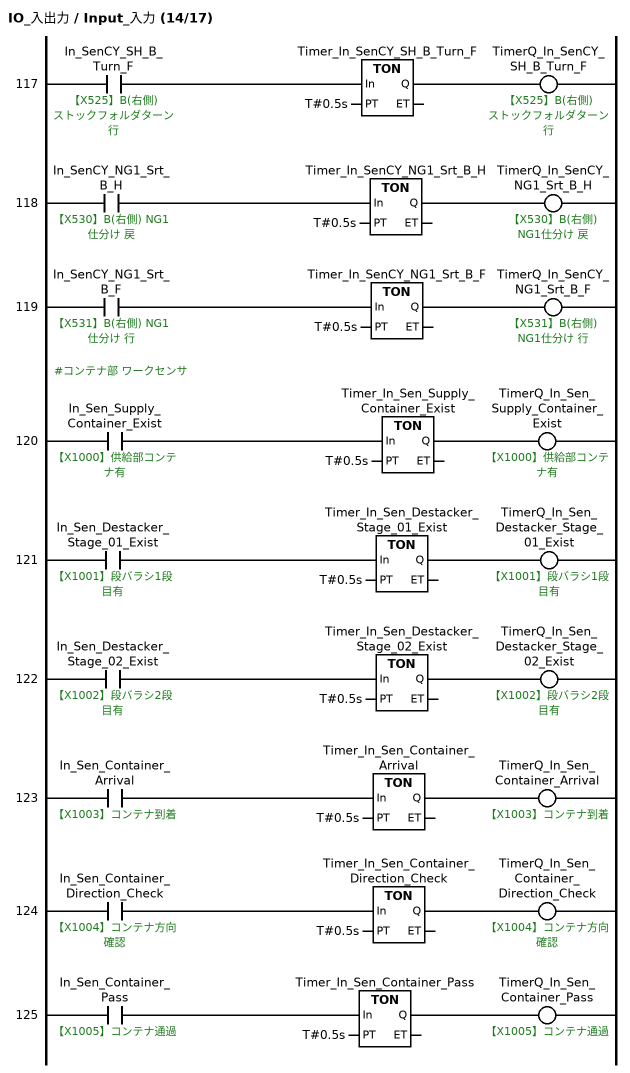
(* [picture p140: IO_入出力 / Input_入力, rungs 117-125] *)
(* Rung 117 *)
Timer_In_SenCY_SH_B_Turn_F(In := In_SenCY_SH_B_Turn_F, PT := T#0.5s);
TimerQ_In_SenCY_SH_B_Turn_F := Timer_In_SenCY_SH_B_Turn_F.Q;
(* Rung 118 *)
Timer_In_SenCY_NG1_Srt_B_H(In := In_SenCY_NG1_Srt_B_H, PT := T#0.5s);
TimerQ_In_SenCY_NG1_Srt_B_H := Timer_In_SenCY_NG1_Srt_B_H.Q;
(* Rung 119 *)
Timer_In_SenCY_NG1_Srt_B_F(In := In_SenCY_NG1_Srt_B_F, PT := T#0.5s);
TimerQ_In_SenCY_NG1_Srt_B_F := Timer_In_SenCY_NG1_Srt_B_F.Q;
(* Rung 120: #コンテナ部 ワークセンサ *)
Timer_In_Sen_Supply_Container_Exist(In := In_Sen_Supply_Container_Exist, PT := T#0.5s);
TimerQ_In_Sen_Supply_Container_Exist := Timer_In_Sen_Supply_Container_Exist.Q;
(* Rung 121 *)
Timer_In_Sen_Destacker_Stage_01_Exist(In := In_Sen_Destacker_Stage_01_Exist, PT := T#0.5s);
TimerQ_In_Sen_Destacker_Stage_01_Exist := Timer_In_Sen_Destacker_Stage_01_Exist.Q;
(* Rung 122 *)
Timer_In_Sen_Destacker_Stage_02_Exist(In := In_Sen_Destacker_Stage_02_Exist, PT := T#0.5s);
TimerQ_In_Sen_Destacker_Stage_02_Exist := Timer_In_Sen_Destacker_Stage_02_Exist.Q;
(* Rung 123 *)
Timer_In_Sen_Container_Arrival(In := In_Sen_Container_Arrival, PT := T#0.5s);
TimerQ_In_Sen_Container_Arrival := Timer_In_Sen_Container_Arrival.Q;
(* Rung 124 *)
Timer_In_Sen_Container_Direction_Check(In := In_Sen_Container_Direction_Check, PT := T#0.5s);
TimerQ_In_Sen_Container_Direction_Check := Timer_In_Sen_Container_Direction_Check.Q;
(* Rung 125 *)
Timer_In_Sen_Container_Pass(In := In_Sen_Container_Pass, PT := T#0.5s);
TimerQ_In_Sen_Container_Pass := Timer_In_Sen_Container_Pass.Q;

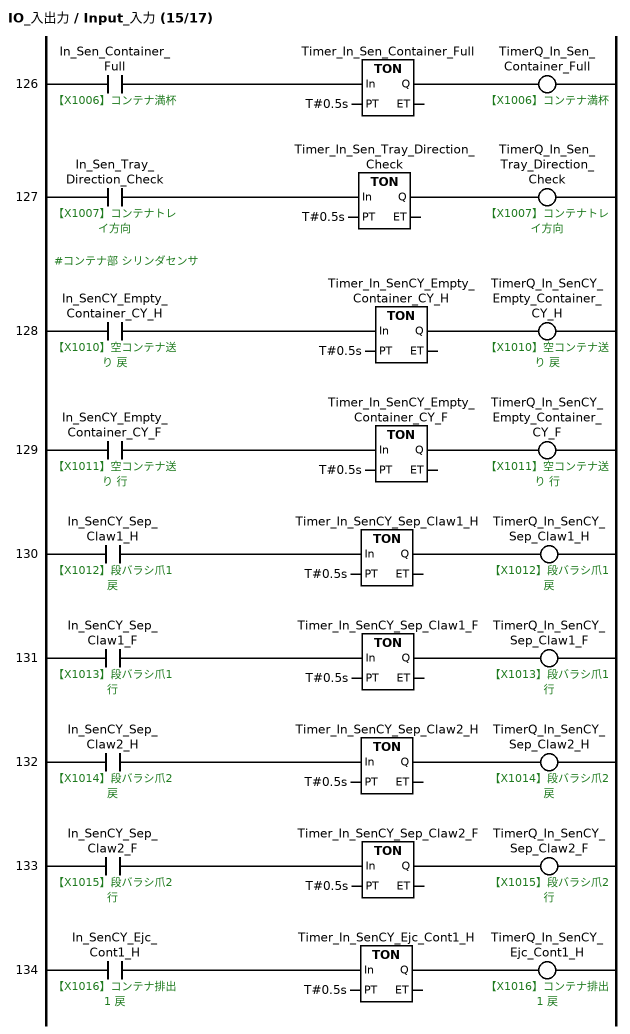
(* Rung 126 *)
Timer_In_Sen_Container_Full(In := In_Sen_Container_Full, PT := T#0.5s);
TimerQ_In_Sen_Container_Full := Timer_In_Sen_Container_Full.Q;
(* Rung 127 *)
Timer_In_Sen_Tray_Direction_Check(In := In_Sen_Tray_Direction_Check, PT := T#0.5s);
TimerQ_In_Sen_Tray_Direction_Check := Timer_In_Sen_Tray_Direction_Check.Q;
(* Rung 128: #コンテナ部 シリンダセンサ *)
Timer_In_SenCY_Empty_Container_CY_H(In := In_SenCY_Empty_Container_CY_H, PT := T#0.5s);
TimerQ_In_SenCY_Empty_Container_CY_H := Timer_In_SenCY_Empty_Container_CY_H.Q;
(* Rung 129 *)
Timer_In_SenCY_Empty_Container_CY_F(In := In_SenCY_Empty_Container_CY_F, PT := T#0.5s);
TimerQ_In_SenCY_Empty_Container_CY_F := Timer_In_SenCY_Empty_Container_CY_F.Q;
(* Rung 130 *)
Timer_In_SenCY_Sep_Claw1_H(In := In_SenCY_Sep_Claw1_H, PT := T#0.5s);
TimerQ_In_SenCY_Sep_Claw1_H := Timer_In_SenCY_Sep_Claw1_H.Q;
(* Rung 131 *)
Timer_In_SenCY_Sep_Claw1_F(In := In_SenCY_Sep_Claw1_F, PT := T#0.5s);
TimerQ_In_SenCY_Sep_Claw1_F := Timer_In_SenCY_Sep_Claw1_F.Q;
(* Rung 132 *)
Timer_In_SenCY_Sep_Claw2_H(In := In_SenCY_Sep_Claw2_H, PT := T#0.5s);
TimerQ_In_SenCY_Sep_Claw2_H := Timer_In_SenCY_Sep_Claw2_H.Q;
(* Rung 133 *)
Timer_In_SenCY_Sep_Claw2_F(In := In_SenCY_Sep_Claw2_F, PT := T#0.5s);
TimerQ_In_SenCY_Sep_Claw2_F := Timer_In_SenCY_Sep_Claw2_F.Q;
(* Rung 134 *)
Timer_In_SenCY_Ejc_Cont1_H(In := In_SenCY_Ejc_Cont1_H, PT := T#0.5s);
TimerQ_In_SenCY_Ejc_Cont1_H := Timer_In_SenCY_Ejc_Cont1_H.Q;

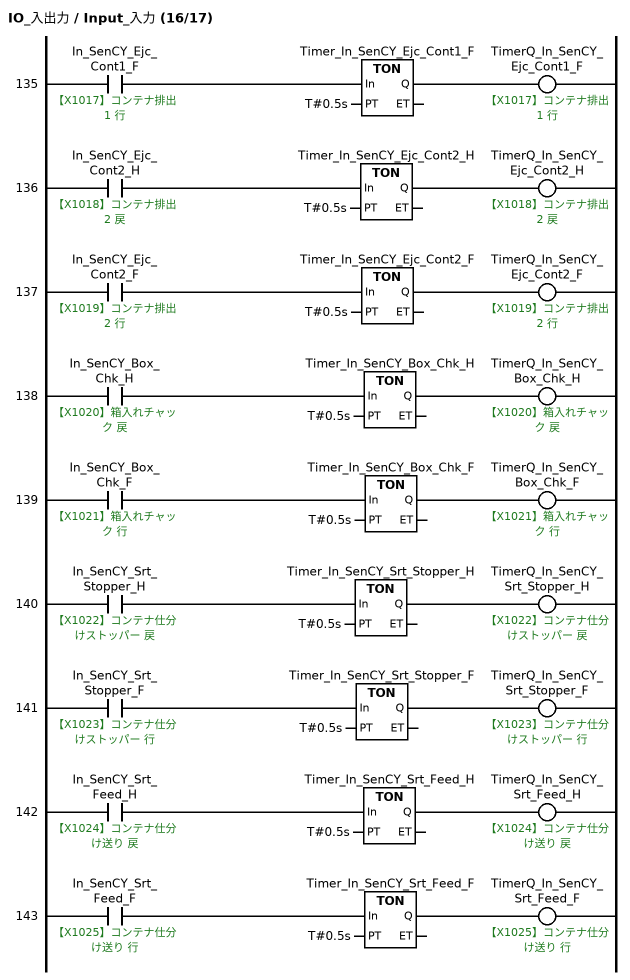
(* Rung 135 *)
Timer_In_SenCY_Ejc_Cont1_F(In := In_SenCY_Ejc_Cont1_F, PT := T#0.5s);
TimerQ_In_SenCY_Ejc_Cont1_F := Timer_In_SenCY_Ejc_Cont1_F.Q;
(* Rung 136 *)
Timer_In_SenCY_Ejc_Cont2_H(In := In_SenCY_Ejc_Cont2_H, PT := T#0.5s);
TimerQ_In_SenCY_Ejc_Cont2_H := Timer_In_SenCY_Ejc_Cont2_H.Q;
(* Rung 137 *)
Timer_In_SenCY_Ejc_Cont2_F(In := In_SenCY_Ejc_Cont2_F, PT := T#0.5s);
TimerQ_In_SenCY_Ejc_Cont2_F := Timer_In_SenCY_Ejc_Cont2_F.Q;
(* Rung 138 *)
Timer_In_SenCY_Box_Chk_H(In := In_SenCY_Box_Chk_H, PT := T#0.5s);
TimerQ_In_SenCY_Box_Chk_H := Timer_In_SenCY_Box_Chk_H.Q;
(* Rung 139 *)
Timer_In_SenCY_Box_Chk_F(In := In_SenCY_Box_Chk_F, PT := T#0.5s);
TimerQ_In_SenCY_Box_Chk_F := Timer_In_SenCY_Box_Chk_F.Q;
(* Rung 140 *)
Timer_In_SenCY_Srt_Stopper_H(In := In_SenCY_Srt_Stopper_H, PT := T#0.5s);
TimerQ_In_SenCY_Srt_Stopper_H := Timer_In_SenCY_Srt_Stopper_H.Q;
(* Rung 141 *)
Timer_In_SenCY_Srt_Stopper_F(In := In_SenCY_Srt_Stopper_F, PT := T#0.5s);
TimerQ_In_SenCY_Srt_Stopper_F := Timer_In_SenCY_Srt_Stopper_F.Q;
(* Rung 142 *)
Timer_In_SenCY_Srt_Feed_H(In := In_SenCY_Srt_Feed_H, PT := T#0.5s);
TimerQ_In_SenCY_Srt_Feed_H := Timer_In_SenCY_Srt_Feed_H.Q;
(* Rung 143 *)
Timer_In_SenCY_Srt_Feed_F(In := In_SenCY_Srt_Feed_F, PT := T#0.5s);
TimerQ_In_SenCY_Srt_Feed_F := Timer_In_SenCY_Srt_Feed_F.Q;

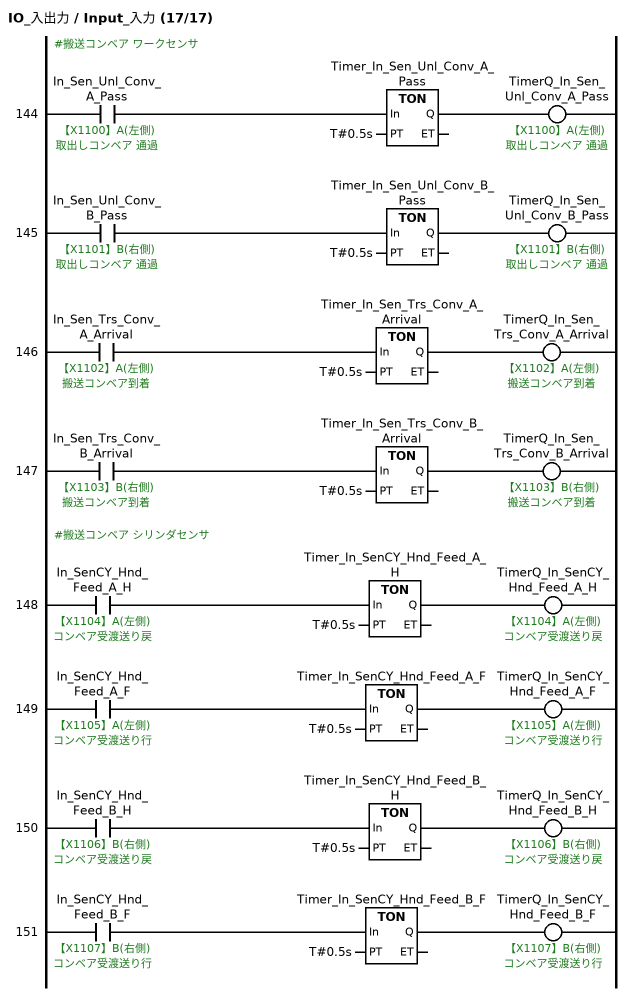
(* Rung 144: #搬送コンベア ワークセンサ *)
Timer_In_Sen_Unl_Conv_A_Pass(In := In_Sen_Unl_Conv_A_Pass, PT := T#0.5s);
TimerQ_In_Sen_Unl_Conv_A_Pass := Timer_In_Sen_Unl_Conv_A_Pass.Q;
(* Rung 145 *)
Timer_In_Sen_Unl_Conv_B_Pass(In := In_Sen_Unl_Conv_B_Pass, PT := T#0.5s);
TimerQ_In_Sen_Unl_Conv_B_Pass := Timer_In_Sen_Unl_Conv_B_Pass.Q;
(* Rung 146 *)
Timer_In_Sen_Trs_Conv_A_Arrival(In := In_Sen_Trs_Conv_A_Arrival, PT := T#0.5s);
TimerQ_In_Sen_Trs_Conv_A_Arrival := Timer_In_Sen_Trs_Conv_A_Arrival.Q;
(* Rung 147 *)
Timer_In_Sen_Trs_Conv_B_Arrival(In := In_Sen_Trs_Conv_B_Arrival, PT := T#0.5s);
TimerQ_In_Sen_Trs_Conv_B_Arrival := Timer_In_Sen_Trs_Conv_B_Arrival.Q;
(* Rung 148: #搬送コンベア シリンダセンサ *)
Timer_In_SenCY_Hnd_Feed_A_H(In := In_SenCY_Hnd_Feed_A_H, PT := T#0.5s);
TimerQ_In_SenCY_Hnd_Feed_A_H := Timer_In_SenCY_Hnd_Feed_A_H.Q;
(* Rung 149 *)
Timer_In_SenCY_Hnd_Feed_A_F(In := In_SenCY_Hnd_Feed_A_F, PT := T#0.5s);
TimerQ_In_SenCY_Hnd_Feed_A_F := Timer_In_SenCY_Hnd_Feed_A_F.Q;
(* Rung 150 *)
Timer_In_SenCY_Hnd_Feed_B_H(In := In_SenCY_Hnd_Feed_B_H, PT := T#0.5s);
TimerQ_In_SenCY_Hnd_Feed_B_H := Timer_In_SenCY_Hnd_Feed_B_H.Q;
(* Rung 151 *)
Timer_In_SenCY_Hnd_Feed_B_F(In := In_SenCY_Hnd_Feed_B_F, PT := T#0.5s);
TimerQ_In_SenCY_Hnd_Feed_B_F := Timer_In_SenCY_Hnd_Feed_B_F.Q;

(* Section Output_出力: ladder, written here as Structured Text *)

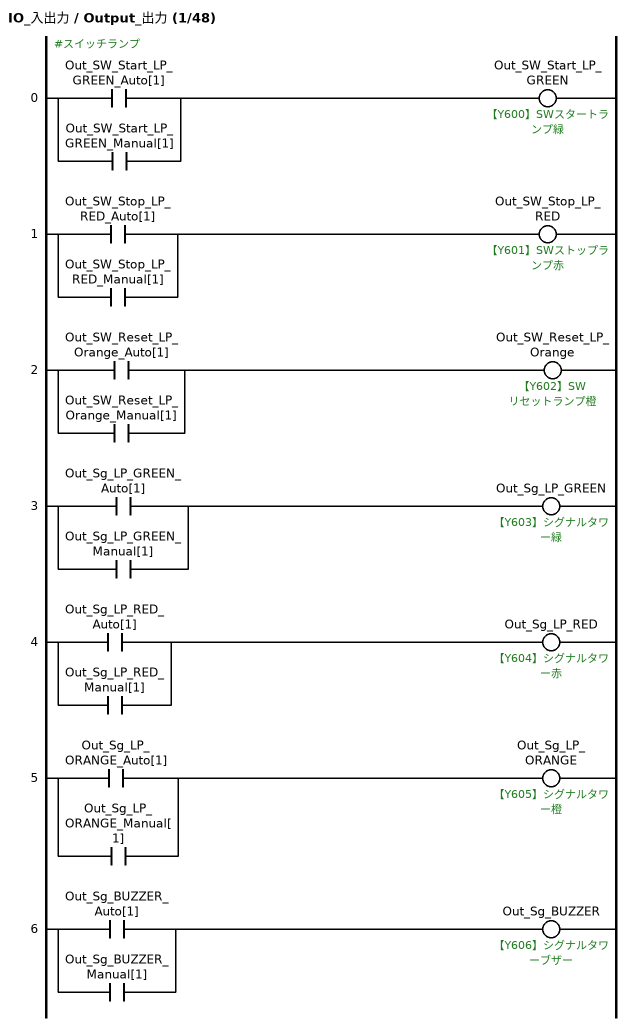
(* Rung 0: #スイッチランプ *)
Out_SW_Start_LP_GREEN := Out_SW_Start_LP_GREEN_Auto[1] OR Out_SW_Start_LP_GREEN_Manual[1];
(* Rung 1 *)
Out_SW_Stop_LP_RED := Out_SW_Stop_LP_RED_Auto[1] OR Out_SW_Stop_LP_RED_Manual[1];
(* Rung 2 *)
Out_SW_Reset_LP_Orange := Out_SW_Reset_LP_Orange_Auto[1] OR Out_SW_Reset_LP_Orange_Manual[1];
(* Rung 3 *)
Out_Sg_LP_GREEN := Out_Sg_LP_GREEN_Auto[1] OR Out_Sg_LP_GREEN_Manual[1];
(* Rung 4 *)
Out_Sg_LP_RED := Out_Sg_LP_RED_Auto[1] OR Out_Sg_LP_RED_Manual[1];
(* Rung 5 *)
Out_Sg_LP_ORANGE := Out_Sg_LP_ORANGE_Auto[1] OR Out_Sg_LP_ORANGE_Manual[1];
(* Rung 6 *)
Out_Sg_BUZZER := Out_Sg_BUZZER_Auto[1] OR Out_Sg_BUZZER_Manual[1];

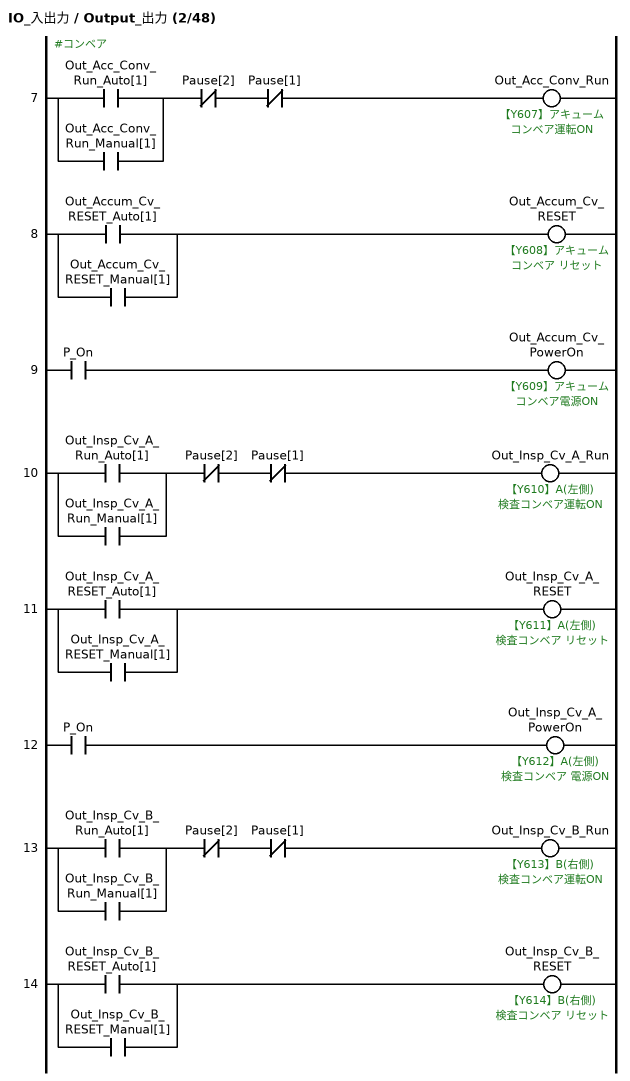
(* Rung 7: #コンベア *)
Out_Acc_Conv_Run := (Out_Acc_Conv_Run_Auto[1] OR Out_Acc_Conv_Run_Manual[1]) AND NOT Pause[2] AND NOT Pause[1];
(* Rung 8 *)
Out_Accum_Cv_RESET := Out_Accum_Cv_RESET_Auto[1] OR Out_Accum_Cv_RESET_Manual[1];
(* Rung 9 *)
Out_Accum_Cv_PowerOn := P_On;
(* Rung 10 *)
Out_Insp_Cv_A_Run := (Out_Insp_Cv_A_Run_Auto[1] OR Out_Insp_Cv_A_Run_Manual[1]) AND NOT Pause[2] AND NOT Pause[1];
(* Rung 11 *)
Out_Insp_Cv_A_RESET := Out_Insp_Cv_A_RESET_Auto[1] OR Out_Insp_Cv_A_RESET_Manual[1];
(* Rung 12 *)
Out_Insp_Cv_A_PowerOn := P_On;
(* Rung 13 *)
Out_Insp_Cv_B_Run := (Out_Insp_Cv_B_Run_Auto[1] OR Out_Insp_Cv_B_Run_Manual[1]) AND NOT Pause[2] AND NOT Pause[1];
(* Rung 14 *)
Out_Insp_Cv_B_RESET := Out_Insp_Cv_B_RESET_Auto[1] OR Out_Insp_Cv_B_RESET_Manual[1];

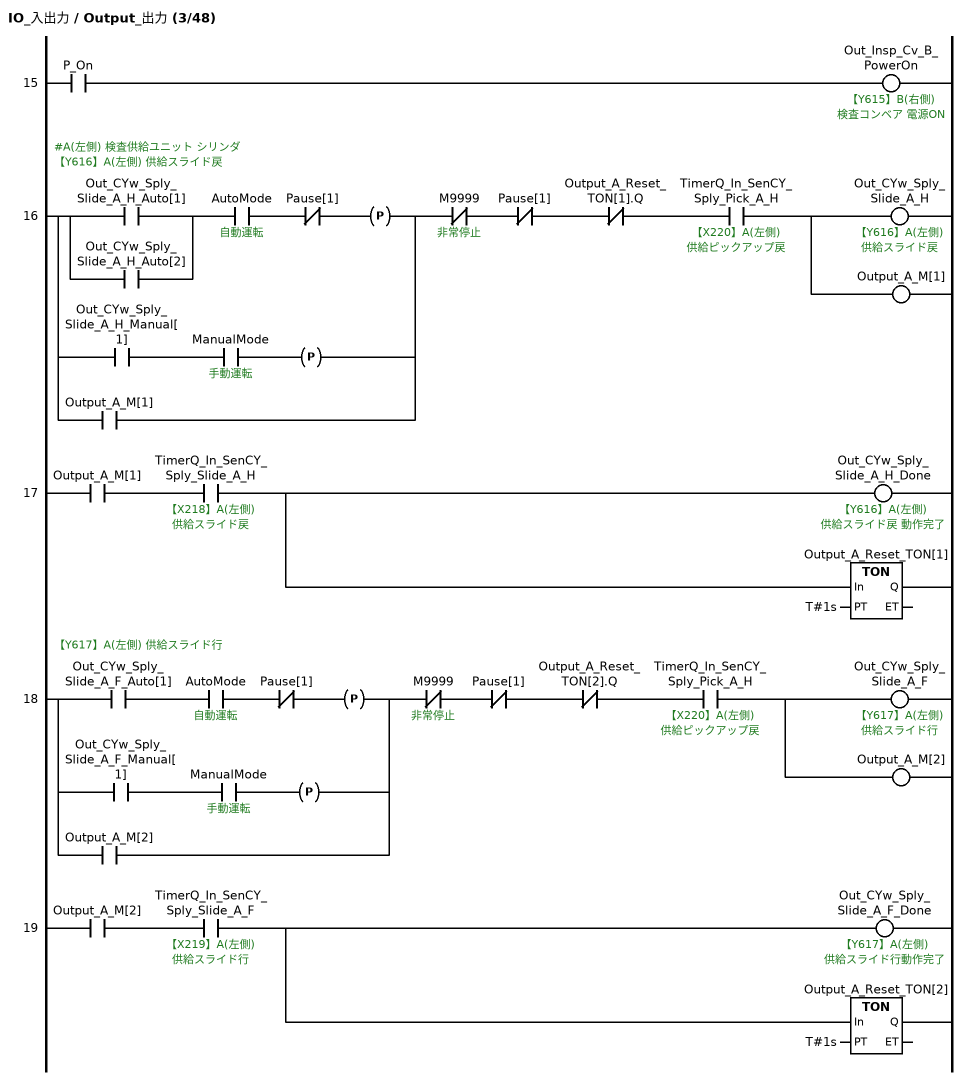
(* Rung 15 *)
Out_Insp_Cv_B_PowerOn := P_On;
(* Rung 16: #A(左側) 検査供給ユニット シリンダ / 【Y616】A(左側) 供給スライド戻 *)
_e1(CLK := (Out_CYw_Sply_Slide_A_H_Auto[1] OR Out_CYw_Sply_Slide_A_H_Auto[2]) AND AutoMode AND NOT Pause[1]);
_e2(CLK := Out_CYw_Sply_Slide_A_H_Manual[1] AND ManualMode);
_p3 := (_e1.Q OR _e2.Q OR Output_A_M[1]) AND NOT M9999 AND NOT Pause[1] AND NOT Output_A_Reset_TON[1].Q AND TimerQ_In_SenCY_Sply_Pick_A_H;
Out_CYw_Sply_Slide_A_H := _p3;
Output_A_M[1] := _p3;
(* Rung 17 *)
Out_CYw_Sply_Slide_A_H_Done := Output_A_M[1] AND TimerQ_In_SenCY_Sply_Slide_A_H;
Output_A_Reset_TON[1](In := Output_A_M[1] AND TimerQ_In_SenCY_Sply_Slide_A_H, PT := T#1s);
(* Rung 18: 【Y617】A(左側) 供給スライド行 *)
_e4(CLK := Out_CYw_Sply_Slide_A_F_Auto[1] AND AutoMode AND NOT Pause[1]);
_e5(CLK := Out_CYw_Sply_Slide_A_F_Manual[1] AND ManualMode);
_p6 := (_e4.Q OR _e5.Q OR Output_A_M[2]) AND NOT M9999 AND NOT Pause[1] AND NOT Output_A_Reset_TON[2].Q AND TimerQ_In_SenCY_Sply_Pick_A_H;
Out_CYw_Sply_Slide_A_F := _p6;
Output_A_M[2] := _p6;
(* Rung 19 *)
Out_CYw_Sply_Slide_A_F_Done := Output_A_M[2] AND TimerQ_In_SenCY_Sply_Slide_A_F;
Output_A_Reset_TON[2](In := Output_A_M[2] AND TimerQ_In_SenCY_Sply_Slide_A_F, PT := T#1s);

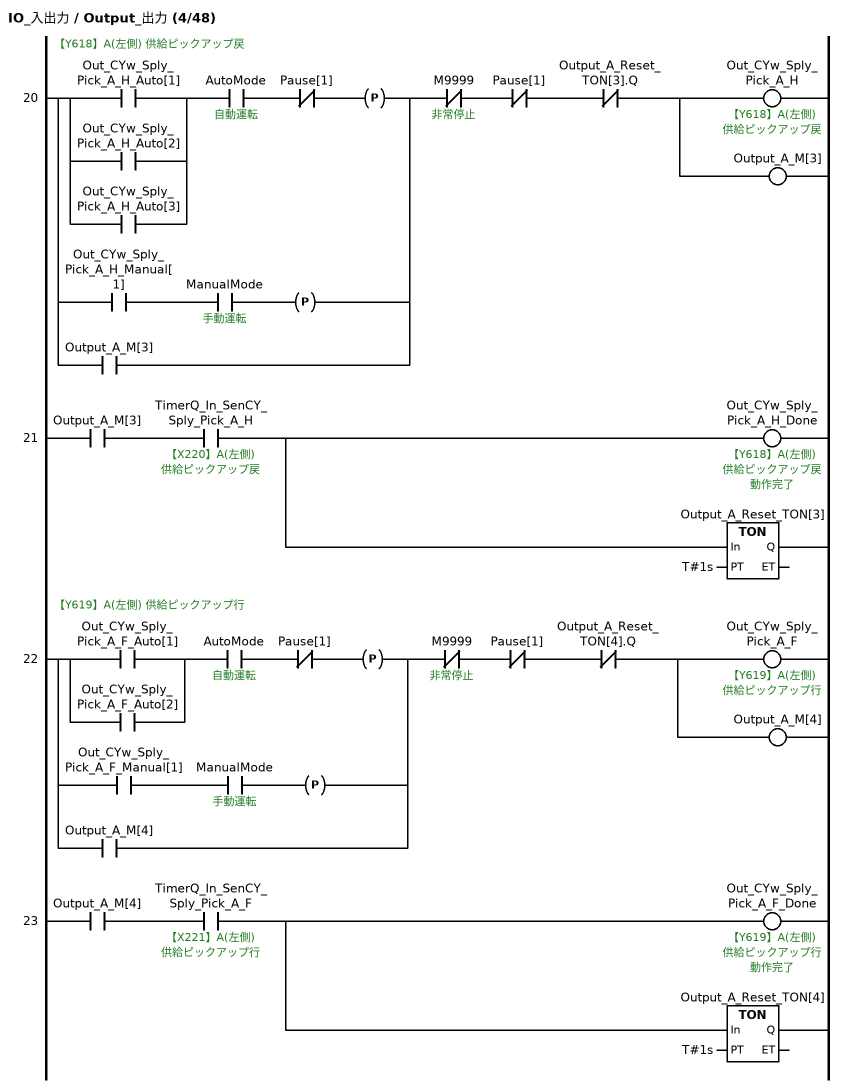
(* Rung 20: 【Y618】A(左側) 供給ピックアップ戻 *)
_e7(CLK := (Out_CYw_Sply_Pick_A_H_Auto[1] OR Out_CYw_Sply_Pick_A_H_Auto[2] OR Out_CYw_Sply_Pick_A_H_Auto[3]) AND AutoMode AND NOT Pause[1]);
_e8(CLK := Out_CYw_Sply_Pick_A_H_Manual[1] AND ManualMode);
_p9 := (_e7.Q OR _e8.Q OR Output_A_M[3]) AND NOT M9999 AND NOT Pause[1] AND NOT Output_A_Reset_TON[3].Q;
Out_CYw_Sply_Pick_A_H := _p9;
Output_A_M[3] := _p9;
(* Rung 21 *)
Out_CYw_Sply_Pick_A_H_Done := Output_A_M[3] AND TimerQ_In_SenCY_Sply_Pick_A_H;
Output_A_Reset_TON[3](In := Output_A_M[3] AND TimerQ_In_SenCY_Sply_Pick_A_H, PT := T#1s);
(* Rung 22: 【Y619】A(左側) 供給ピックアップ行 *)
_e10(CLK := (Out_CYw_Sply_Pick_A_F_Auto[1] OR Out_CYw_Sply_Pick_A_F_Auto[2]) AND AutoMode AND NOT Pause[1]);
_e11(CLK := Out_CYw_Sply_Pick_A_F_Manual[1] AND ManualMode);
_p12 := (_e10.Q OR _e11.Q OR Output_A_M[4]) AND NOT M9999 AND NOT Pause[1] AND NOT Output_A_Reset_TON[4].Q;
Out_CYw_Sply_Pick_A_F := _p12;
Output_A_M[4] := _p12;
(* Rung 23 *)
Out_CYw_Sply_Pick_A_F_Done := Output_A_M[4] AND TimerQ_In_SenCY_Sply_Pick_A_F;
Output_A_Reset_TON[4](In := Output_A_M[4] AND TimerQ_In_SenCY_Sply_Pick_A_F, PT := T#1s);

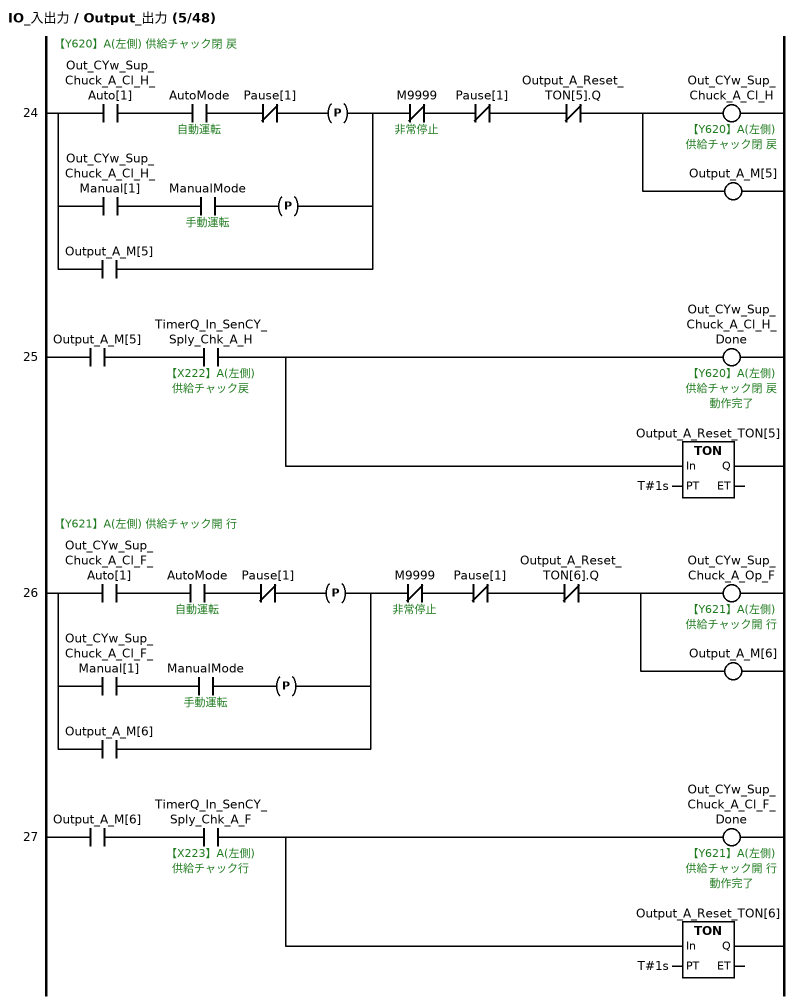
(* Rung 24: 【Y620】A(左側) 供給チャック閉 戻 *)
_e13(CLK := Out_CYw_Sup_Chuck_A_Cl_H_Auto[1] AND AutoMode AND NOT Pause[1]);
_e14(CLK := Out_CYw_Sup_Chuck_A_Cl_H_Manual[1] AND ManualMode);
_p15 := (_e13.Q OR _e14.Q OR Output_A_M[5]) AND NOT M9999 AND NOT Pause[1] AND NOT Output_A_Reset_TON[5].Q;
Out_CYw_Sup_Chuck_A_Cl_H := _p15;
Output_A_M[5] := _p15;
(* Rung 25 *)
Out_CYw_Sup_Chuck_A_Cl_H_Done := Output_A_M[5] AND TimerQ_In_SenCY_Sply_Chk_A_H;
Output_A_Reset_TON[5](In := Output_A_M[5] AND TimerQ_In_SenCY_Sply_Chk_A_H, PT := T#1s);
(* Rung 26: 【Y621】A(左側) 供給チャック開 行 *)
_e16(CLK := Out_CYw_Sup_Chuck_A_Cl_F_Auto[1] AND AutoMode AND NOT Pause[1]);
_e17(CLK := Out_CYw_Sup_Chuck_A_Cl_F_Manual[1] AND ManualMode);
_p18 := (_e16.Q OR _e17.Q OR Output_A_M[6]) AND NOT M9999 AND NOT Pause[1] AND NOT Output_A_Reset_TON[6].Q;
Out_CYw_Sup_Chuck_A_Op_F := _p18;
Output_A_M[6] := _p18;
(* Rung 27 *)
Out_CYw_Sup_Chuck_A_Cl_F_Done := Output_A_M[6] AND TimerQ_In_SenCY_Sply_Chk_A_F;
Output_A_Reset_TON[6](In := Output_A_M[6] AND TimerQ_In_SenCY_Sply_Chk_A_F, PT := T#1s);

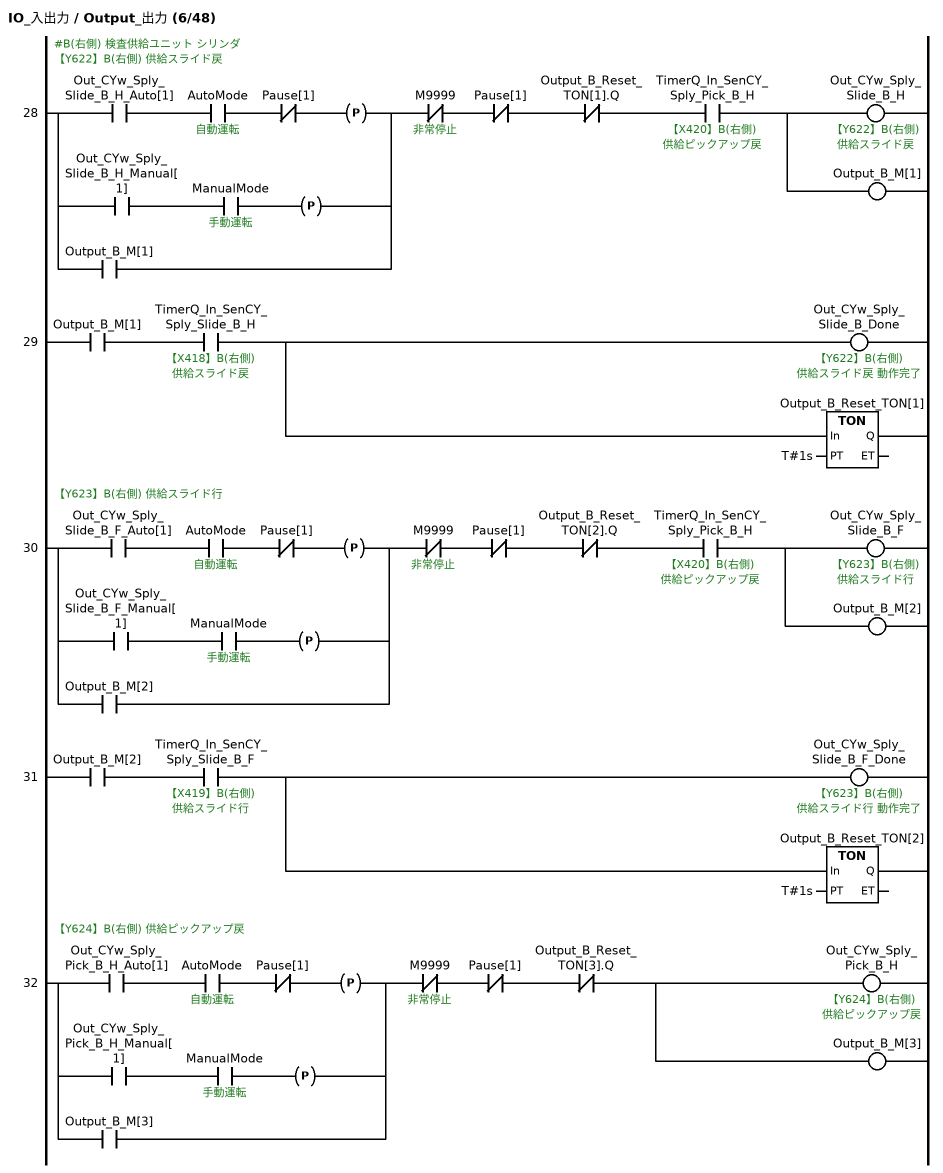
(* Rung 28: #B(右側) 検査供給ユニット シリンダ / 【Y622】B(右側) 供給スライド戻 *)
_e19(CLK := Out_CYw_Sply_Slide_B_H_Auto[1] AND AutoMode AND NOT Pause[1]);
_e20(CLK := Out_CYw_Sply_Slide_B_H_Manual[1] AND ManualMode);
_p21 := (_e19.Q OR _e20.Q OR Output_B_M[1]) AND NOT M9999 AND NOT Pause[1] AND NOT Output_B_Reset_TON[1].Q AND TimerQ_In_SenCY_Sply_Pick_B_H;
Out_CYw_Sply_Slide_B_H := _p21;
Output_B_M[1] := _p21;
(* Rung 29 *)
Out_CYw_Sply_Slide_B_Done := Output_B_M[1] AND TimerQ_In_SenCY_Sply_Slide_B_H;
Output_B_Reset_TON[1](In := Output_B_M[1] AND TimerQ_In_SenCY_Sply_Slide_B_H, PT := T#1s);
(* Rung 30: 【Y623】B(右側) 供給スライド行 *)
_e22(CLK := Out_CYw_Sply_Slide_B_F_Auto[1] AND AutoMode AND NOT Pause[1]);
_e23(CLK := Out_CYw_Sply_Slide_B_F_Manual[1] AND ManualMode);
_p24 := (_e22.Q OR _e23.Q OR Output_B_M[2]) AND NOT M9999 AND NOT Pause[1] AND NOT Output_B_Reset_TON[2].Q AND TimerQ_In_SenCY_Sply_Pick_B_H;
Out_CYw_Sply_Slide_B_F := _p24;
Output_B_M[2] := _p24;
(* Rung 31 *)
Out_CYw_Sply_Slide_B_F_Done := Output_B_M[2] AND TimerQ_In_SenCY_Sply_Slide_B_F;
Output_B_Reset_TON[2](In := Output_B_M[2] AND TimerQ_In_SenCY_Sply_Slide_B_F, PT := T#1s);
(* Rung 32: 【Y624】B(右側) 供給ピックアップ戻 *)
_e25(CLK := Out_CYw_Sply_Pick_B_H_Auto[1] AND AutoMode AND NOT Pause[1]);
_e26(CLK := Out_CYw_Sply_Pick_B_H_Manual[1] AND ManualMode);
_p27 := (_e25.Q OR _e26.Q OR Output_B_M[3]) AND NOT M9999 AND NOT Pause[1] AND NOT Output_B_Reset_TON[3].Q;
Out_CYw_Sply_Pick_B_H := _p27;
Output_B_M[3] := _p27;

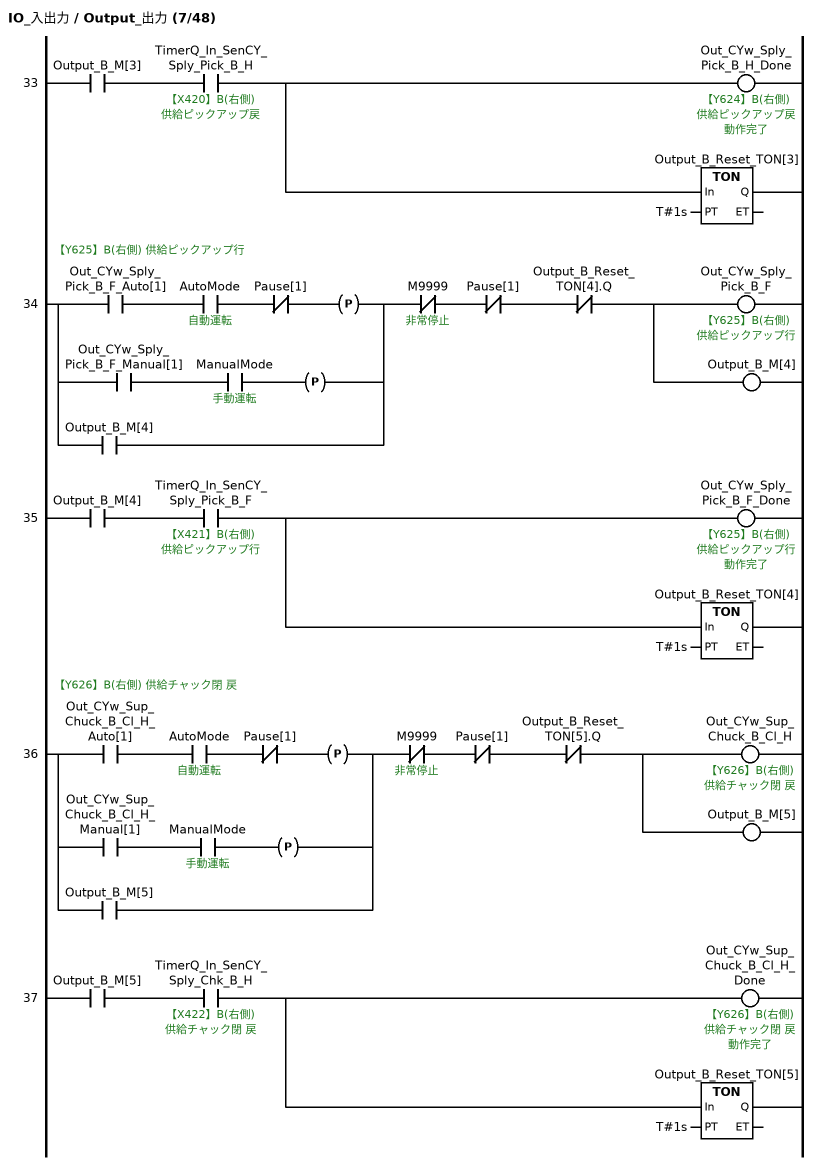
(* Rung 33 *)
Out_CYw_Sply_Pick_B_H_Done := Output_B_M[3] AND TimerQ_In_SenCY_Sply_Pick_B_H;
Output_B_Reset_TON[3](In := Output_B_M[3] AND TimerQ_In_SenCY_Sply_Pick_B_H, PT := T#1s);
(* Rung 34: 【Y625】B(右側) 供給ピックアップ行 *)
_e28(CLK := Out_CYw_Sply_Pick_B_F_Auto[1] AND AutoMode AND NOT Pause[1]);
_e29(CLK := Out_CYw_Sply_Pick_B_F_Manual[1] AND ManualMode);
_p30 := (_e28.Q OR _e29.Q OR Output_B_M[4]) AND NOT M9999 AND NOT Pause[1] AND NOT Output_B_Reset_TON[4].Q;
Out_CYw_Sply_Pick_B_F := _p30;
Output_B_M[4] := _p30;
(* Rung 35 *)
Out_CYw_Sply_Pick_B_F_Done := Output_B_M[4] AND TimerQ_In_SenCY_Sply_Pick_B_F;
Output_B_Reset_TON[4](In := Output_B_M[4] AND TimerQ_In_SenCY_Sply_Pick_B_F, PT := T#1s);
(* Rung 36: 【Y626】B(右側) 供給チャック閉 戻 *)
_e31(CLK := Out_CYw_Sup_Chuck_B_Cl_H_Auto[1] AND AutoMode AND NOT Pause[1]);
_e32(CLK := Out_CYw_Sup_Chuck_B_Cl_H_Manual[1] AND ManualMode);
_p33 := (_e31.Q OR _e32.Q OR Output_B_M[5]) AND NOT M9999 AND NOT Pause[1] AND NOT Output_B_Reset_TON[5].Q;
Out_CYw_Sup_Chuck_B_Cl_H := _p33;
Output_B_M[5] := _p33;
(* Rung 37 *)
Out_CYw_Sup_Chuck_B_Cl_H_Done := Output_B_M[5] AND TimerQ_In_SenCY_Sply_Chk_B_H;
Output_B_Reset_TON[5](In := Output_B_M[5] AND TimerQ_In_SenCY_Sply_Chk_B_H, PT := T#1s);

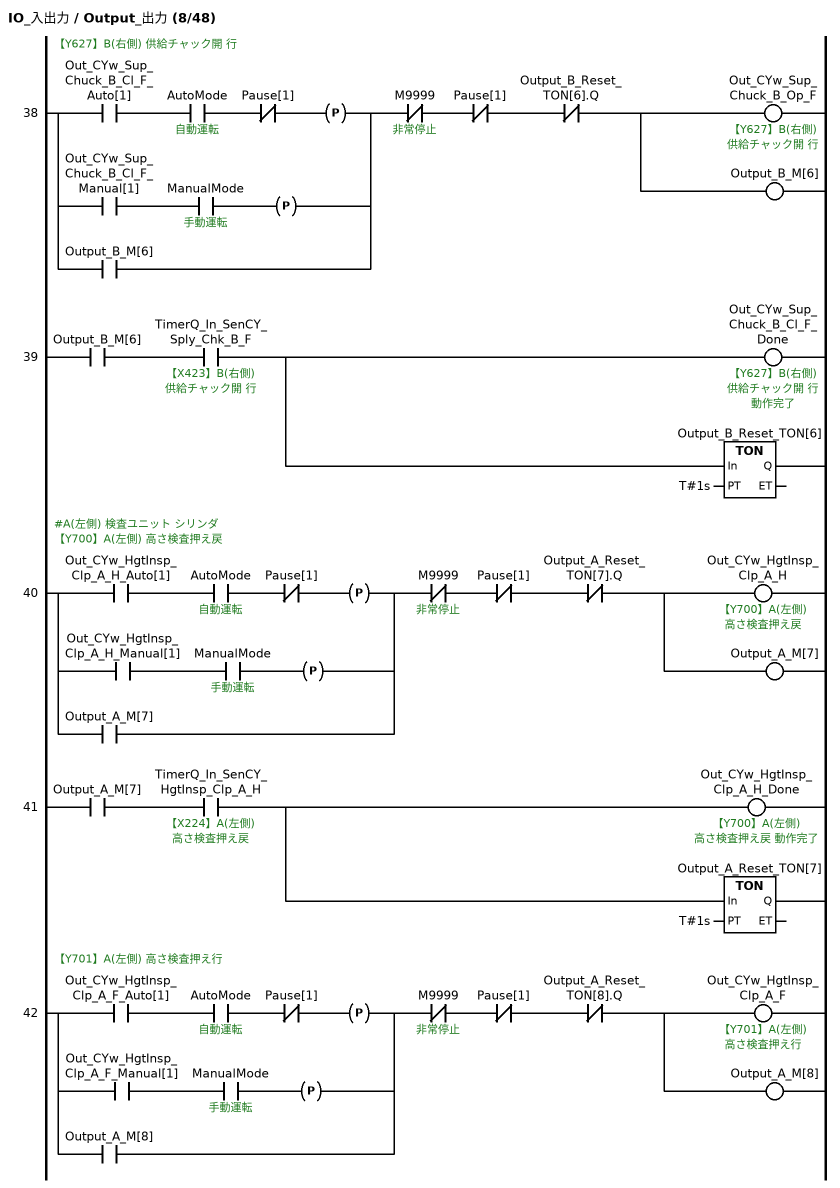
(* Rung 38: 【Y627】B(右側) 供給チャック開 行 *)
_e34(CLK := Out_CYw_Sup_Chuck_B_Cl_F_Auto[1] AND AutoMode AND NOT Pause[1]);
_e35(CLK := Out_CYw_Sup_Chuck_B_Cl_F_Manual[1] AND ManualMode);
_p36 := (_e34.Q OR _e35.Q OR Output_B_M[6]) AND NOT M9999 AND NOT Pause[1] AND NOT Output_B_Reset_TON[6].Q;
Out_CYw_Sup_Chuck_B_Op_F := _p36;
Output_B_M[6] := _p36;
(* Rung 39 *)
Out_CYw_Sup_Chuck_B_Cl_F_Done := Output_B_M[6] AND TimerQ_In_SenCY_Sply_Chk_B_F;
Output_B_Reset_TON[6](In := Output_B_M[6] AND TimerQ_In_SenCY_Sply_Chk_B_F, PT := T#1s);
(* Rung 40: #A(左側) 検査ユニット シリンダ / 【Y700】A(左側) 高さ検査押え戻 *)
_e37(CLK := Out_CYw_HgtInsp_Clp_A_H_Auto[1] AND AutoMode AND NOT Pause[1]);
_e38(CLK := Out_CYw_HgtInsp_Clp_A_H_Manual[1] AND ManualMode);
_p39 := (_e37.Q OR _e38.Q OR Output_A_M[7]) AND NOT M9999 AND NOT Pause[1] AND NOT Output_A_Reset_TON[7].Q;
Out_CYw_HgtInsp_Clp_A_H := _p39;
Output_A_M[7] := _p39;
(* Rung 41 *)
_p40 := Output_A_M[7] AND TimerQ_In_SenCY_HgtInsp_Clp_A_H;
Out_CYw_HgtInsp_Clp_A_H_Done := _p40;
Output_A_Reset_TON[7](In := _p40, PT := T#1s);
(* Rung 42: 【Y701】A(左側) 高さ検査押え行 *)
_e41(CLK := Out_CYw_HgtInsp_Clp_A_F_Auto[1] AND AutoMode AND NOT Pause[1]);
_e42(CLK := Out_CYw_HgtInsp_Clp_A_F_Manual[1] AND ManualMode);
_p43 := (_e41.Q OR _e42.Q OR Output_A_M[8]) AND NOT M9999 AND NOT Pause[1] AND NOT Output_A_Reset_TON[8].Q;
Out_CYw_HgtInsp_Clp_A_F := _p43;
Output_A_M[8] := _p43;

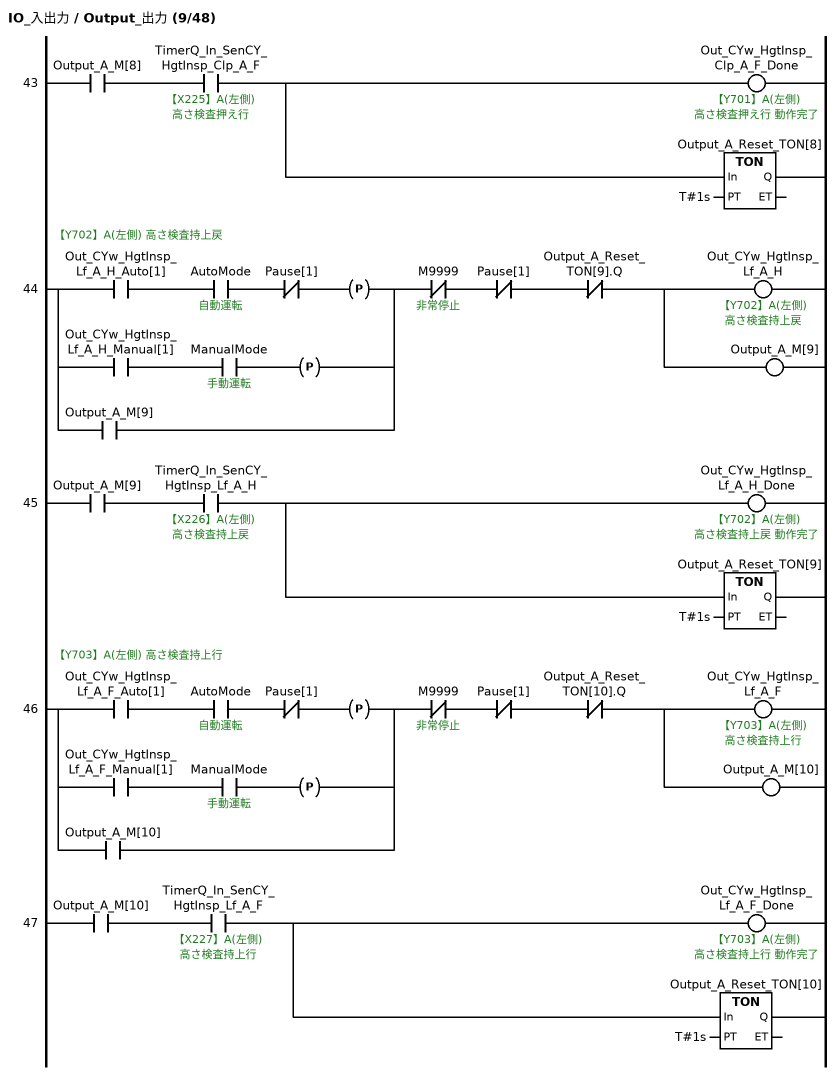
(* Rung 43 *)
_p44 := Output_A_M[8] AND TimerQ_In_SenCY_HgtInsp_Clp_A_F;
Out_CYw_HgtInsp_Clp_A_F_Done := _p44;
Output_A_Reset_TON[8](In := _p44, PT := T#1s);
(* Rung 44: 【Y702】A(左側) 高さ検査持上戻 *)
_e45(CLK := Out_CYw_HgtInsp_Lf_A_H_Auto[1] AND AutoMode AND NOT Pause[1]);
_e46(CLK := Out_CYw_HgtInsp_Lf_A_H_Manual[1] AND ManualMode);
_p47 := (_e45.Q OR _e46.Q OR Output_A_M[9]) AND NOT M9999 AND NOT Pause[1] AND NOT Output_A_Reset_TON[9].Q;
Out_CYw_HgtInsp_Lf_A_H := _p47;
Output_A_M[9] := _p47;
(* Rung 45 *)
Out_CYw_HgtInsp_Lf_A_H_Done := Output_A_M[9] AND TimerQ_In_SenCY_HgtInsp_Lf_A_H;
Output_A_Reset_TON[9](In := Output_A_M[9] AND TimerQ_In_SenCY_HgtInsp_Lf_A_H, PT := T#1s);
(* Rung 46: 【Y703】A(左側) 高さ検査持上行 *)
_e48(CLK := Out_CYw_HgtInsp_Lf_A_F_Auto[1] AND AutoMode AND NOT Pause[1]);
_e49(CLK := Out_CYw_HgtInsp_Lf_A_F_Manual[1] AND ManualMode);
_p50 := (_e48.Q OR _e49.Q OR Output_A_M[10]) AND NOT M9999 AND NOT Pause[1] AND NOT Output_A_Reset_TON[10].Q;
Out_CYw_HgtInsp_Lf_A_F := _p50;
Output_A_M[10] := _p50;
(* Rung 47 *)
_p51 := Output_A_M[10] AND TimerQ_In_SenCY_HgtInsp_Lf_A_F;
Out_CYw_HgtInsp_Lf_A_F_Done := _p51;
Output_A_Reset_TON[10](In := _p51, PT := T#1s);

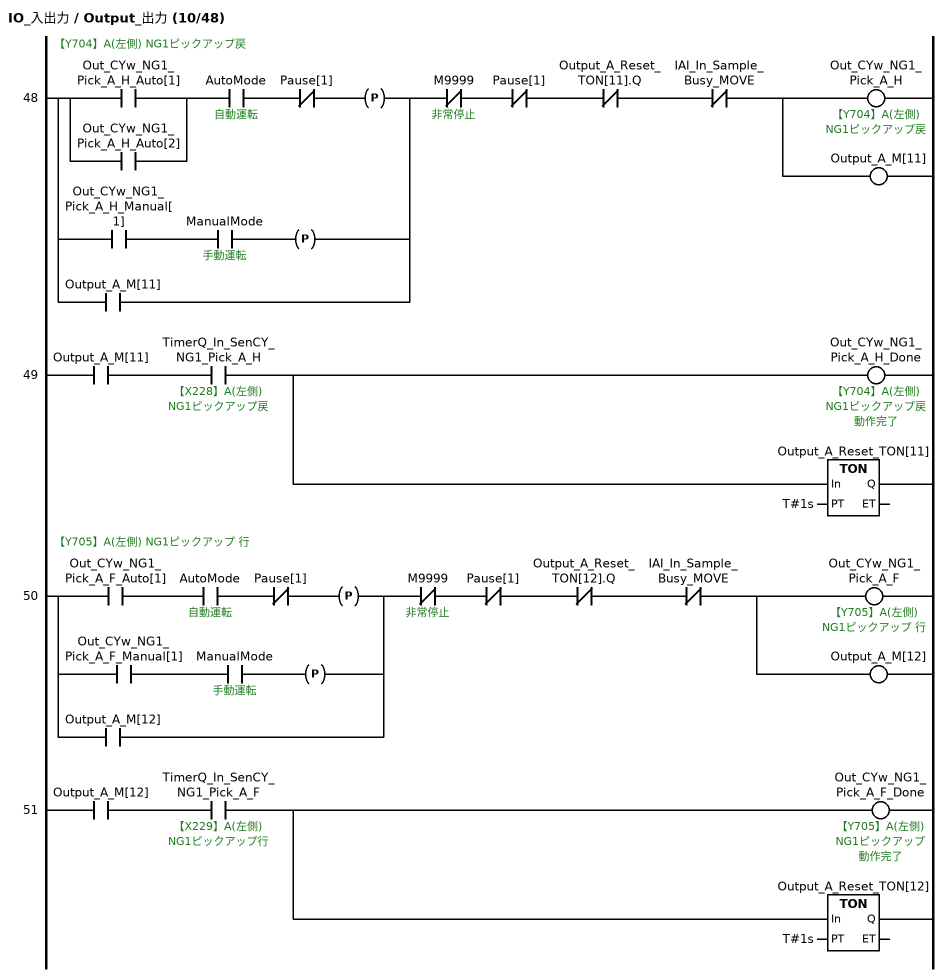
(* Rung 48: 【Y704】A(左側) NG1ピックアップ戻 *)
_e52(CLK := (Out_CYw_NG1_Pick_A_H_Auto[1] OR Out_CYw_NG1_Pick_A_H_Auto[2]) AND AutoMode AND NOT Pause[1]);
_e53(CLK := Out_CYw_NG1_Pick_A_H_Manual[1] AND ManualMode);
_p54 := (_e52.Q OR _e53.Q OR Output_A_M[11]) AND NOT M9999 AND NOT Pause[1] AND NOT Output_A_Reset_TON[11].Q AND NOT IAI_In_Sample_Busy_MOVE;
Out_CYw_NG1_Pick_A_H := _p54;
Output_A_M[11] := _p54;
(* Rung 49 *)
Out_CYw_NG1_Pick_A_H_Done := Output_A_M[11] AND TimerQ_In_SenCY_NG1_Pick_A_H;
Output_A_Reset_TON[11](In := Output_A_M[11] AND TimerQ_In_SenCY_NG1_Pick_A_H, PT := T#1s);
(* Rung 50: 【Y705】A(左側) NG1ピックアップ 行 *)
_e55(CLK := Out_CYw_NG1_Pick_A_F_Auto[1] AND AutoMode AND NOT Pause[1]);
_e56(CLK := Out_CYw_NG1_Pick_A_F_Manual[1] AND ManualMode);
_p57 := (_e55.Q OR _e56.Q OR Output_A_M[12]) AND NOT M9999 AND NOT Pause[1] AND NOT Output_A_Reset_TON[12].Q AND NOT IAI_In_Sample_Busy_MOVE;
Out_CYw_NG1_Pick_A_F := _p57;
Output_A_M[12] := _p57;
(* Rung 51 *)
Out_CYw_NG1_Pick_A_F_Done := Output_A_M[12] AND TimerQ_In_SenCY_NG1_Pick_A_F;
Output_A_Reset_TON[12](In := Output_A_M[12] AND TimerQ_In_SenCY_NG1_Pick_A_F, PT := T#1s);

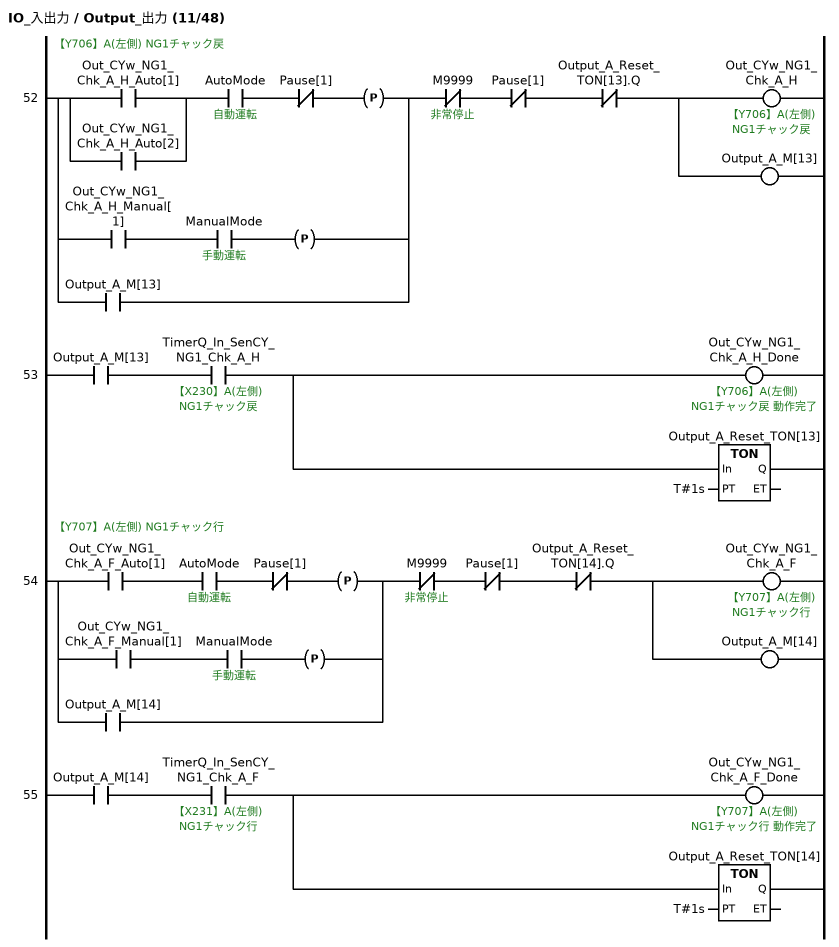
(* Rung 52: 【Y706】A(左側) NG1チャック戻 *)
_e58(CLK := (Out_CYw_NG1_Chk_A_H_Auto[1] OR Out_CYw_NG1_Chk_A_H_Auto[2]) AND AutoMode AND NOT Pause[1]);
_e59(CLK := Out_CYw_NG1_Chk_A_H_Manual[1] AND ManualMode);
_p60 := (_e58.Q OR _e59.Q OR Output_A_M[13]) AND NOT M9999 AND NOT Pause[1] AND NOT Output_A_Reset_TON[13].Q;
Out_CYw_NG1_Chk_A_H := _p60;
Output_A_M[13] := _p60;
(* Rung 53 *)
Out_CYw_NG1_Chk_A_H_Done := Output_A_M[13] AND TimerQ_In_SenCY_NG1_Chk_A_H;
Output_A_Reset_TON[13](In := Output_A_M[13] AND TimerQ_In_SenCY_NG1_Chk_A_H, PT := T#1s);
(* Rung 54: 【Y707】A(左側) NG1チャック行 *)
_e61(CLK := Out_CYw_NG1_Chk_A_F_Auto[1] AND AutoMode AND NOT Pause[1]);
_e62(CLK := Out_CYw_NG1_Chk_A_F_Manual[1] AND ManualMode);
_p63 := (_e61.Q OR _e62.Q OR Output_A_M[14]) AND NOT M9999 AND NOT Pause[1] AND NOT Output_A_Reset_TON[14].Q;
Out_CYw_NG1_Chk_A_F := _p63;
Output_A_M[14] := _p63;
(* Rung 55 *)
Out_CYw_NG1_Chk_A_F_Done := Output_A_M[14] AND TimerQ_In_SenCY_NG1_Chk_A_F;
Output_A_Reset_TON[14](In := Output_A_M[14] AND TimerQ_In_SenCY_NG1_Chk_A_F, PT := T#1s);

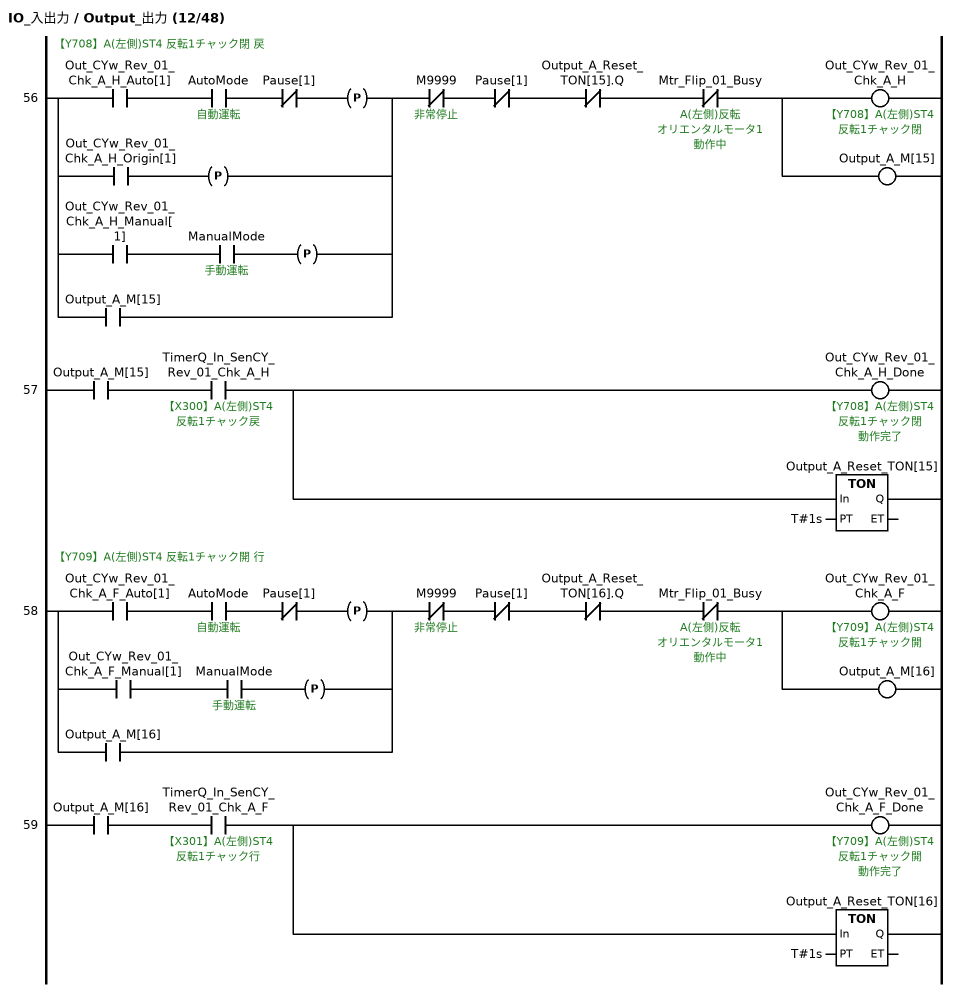
(* Rung 56: 【Y708】A(左側)ST4 反転1チャック閉 戻 *)
_e64(CLK := Out_CYw_Rev_01_Chk_A_H_Auto[1] AND AutoMode AND NOT Pause[1]);
_e65(CLK := Out_CYw_Rev_01_Chk_A_H_Origin[1]);
_e66(CLK := Out_CYw_Rev_01_Chk_A_H_Manual[1] AND ManualMode);
_p67 := (_e64.Q OR _e65.Q OR _e66.Q OR Output_A_M[15]) AND NOT M9999 AND NOT Pause[1] AND NOT Output_A_Reset_TON[15].Q AND NOT Mtr_Flip_01_Busy;
Out_CYw_Rev_01_Chk_A_H := _p67;
Output_A_M[15] := _p67;
(* Rung 57 *)
_p68 := Output_A_M[15] AND TimerQ_In_SenCY_Rev_01_Chk_A_H;
Out_CYw_Rev_01_Chk_A_H_Done := _p68;
Output_A_Reset_TON[15](In := _p68, PT := T#1s);
(* Rung 58: 【Y709】A(左側)ST4 反転1チャック開 行 *)
_e69(CLK := Out_CYw_Rev_01_Chk_A_F_Auto[1] AND AutoMode AND NOT Pause[1]);
_e70(CLK := Out_CYw_Rev_01_Chk_A_F_Manual[1] AND ManualMode);
_p71 := (_e69.Q OR _e70.Q OR Output_A_M[16]) AND NOT M9999 AND NOT Pause[1] AND NOT Output_A_Reset_TON[16].Q AND NOT Mtr_Flip_01_Busy;
Out_CYw_Rev_01_Chk_A_F := _p71;
Output_A_M[16] := _p71;
(* Rung 59 *)
_p72 := Output_A_M[16] AND TimerQ_In_SenCY_Rev_01_Chk_A_F;
Out_CYw_Rev_01_Chk_A_F_Done := _p72;
Output_A_Reset_TON[16](In := _p72, PT := T#1s);

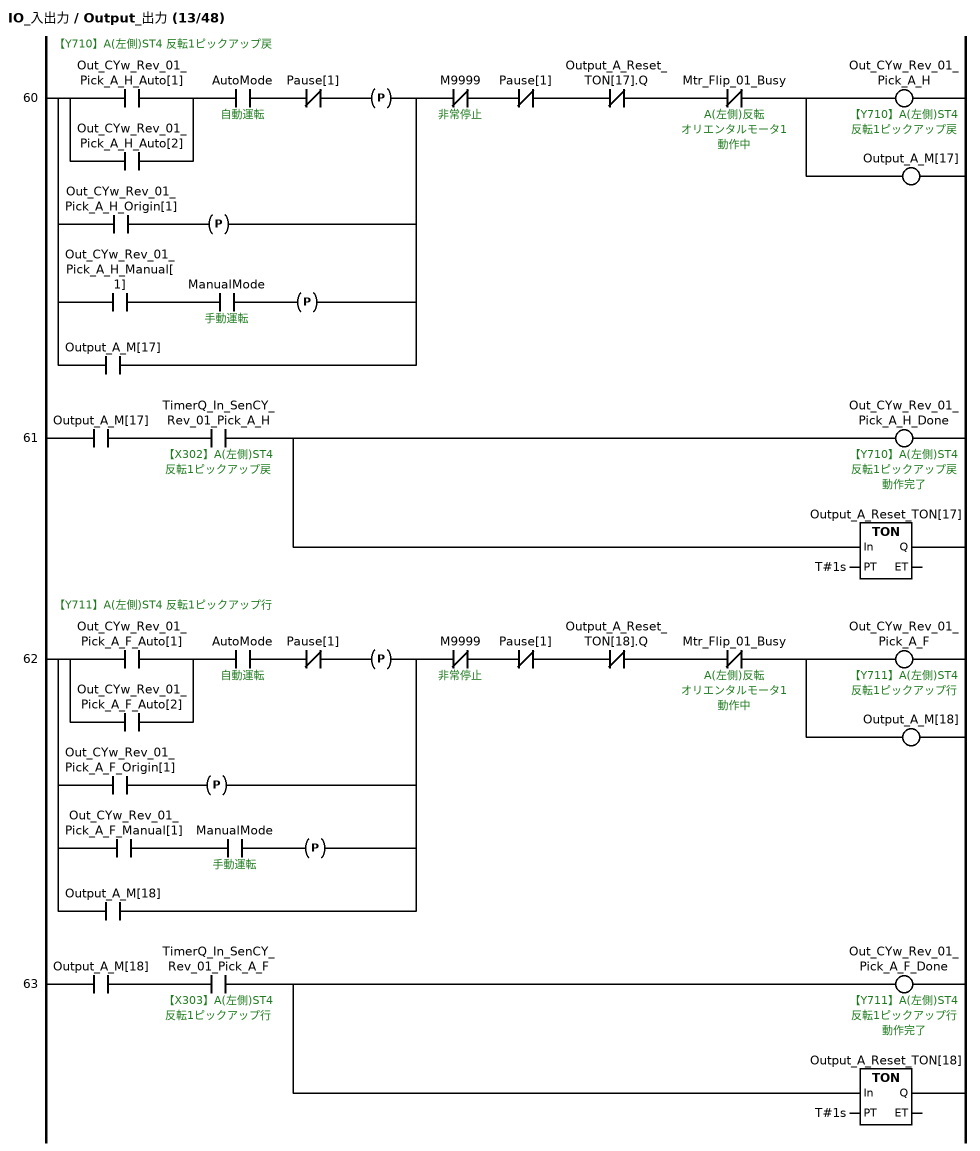
(* Rung 60: 【Y710】A(左側)ST4 反転1ピックアップ戻 *)
_e73(CLK := (Out_CYw_Rev_01_Pick_A_H_Auto[1] OR Out_CYw_Rev_01_Pick_A_H_Auto[2]) AND AutoMode AND NOT Pause[1]);
_e74(CLK := Out_CYw_Rev_01_Pick_A_H_Origin[1]);
_e75(CLK := Out_CYw_Rev_01_Pick_A_H_Manual[1] AND ManualMode);
_p76 := (_e73.Q OR _e74.Q OR _e75.Q OR Output_A_M[17]) AND NOT M9999 AND NOT Pause[1] AND NOT Output_A_Reset_TON[17].Q AND NOT Mtr_Flip_01_Busy;
Out_CYw_Rev_01_Pick_A_H := _p76;
Output_A_M[17] := _p76;
(* Rung 61 *)
_p77 := Output_A_M[17] AND TimerQ_In_SenCY_Rev_01_Pick_A_H;
Out_CYw_Rev_01_Pick_A_H_Done := _p77;
Output_A_Reset_TON[17](In := _p77, PT := T#1s);
(* Rung 62: 【Y711】A(左側)ST4 反転1ピックアップ行 *)
_e78(CLK := (Out_CYw_Rev_01_Pick_A_F_Auto[1] OR Out_CYw_Rev_01_Pick_A_F_Auto[2]) AND AutoMode AND NOT Pause[1]);
_e79(CLK := Out_CYw_Rev_01_Pick_A_F_Origin[1]);
_e80(CLK := Out_CYw_Rev_01_Pick_A_F_Manual[1] AND ManualMode);
_p81 := (_e78.Q OR _e79.Q OR _e80.Q OR Output_A_M[18]) AND NOT M9999 AND NOT Pause[1] AND NOT Output_A_Reset_TON[18].Q AND NOT Mtr_Flip_01_Busy;
Out_CYw_Rev_01_Pick_A_F := _p81;
Output_A_M[18] := _p81;
(* Rung 63 *)
_p82 := Output_A_M[18] AND TimerQ_In_SenCY_Rev_01_Pick_A_F;
Out_CYw_Rev_01_Pick_A_F_Done := _p82;
Output_A_Reset_TON[18](In := _p82, PT := T#1s);

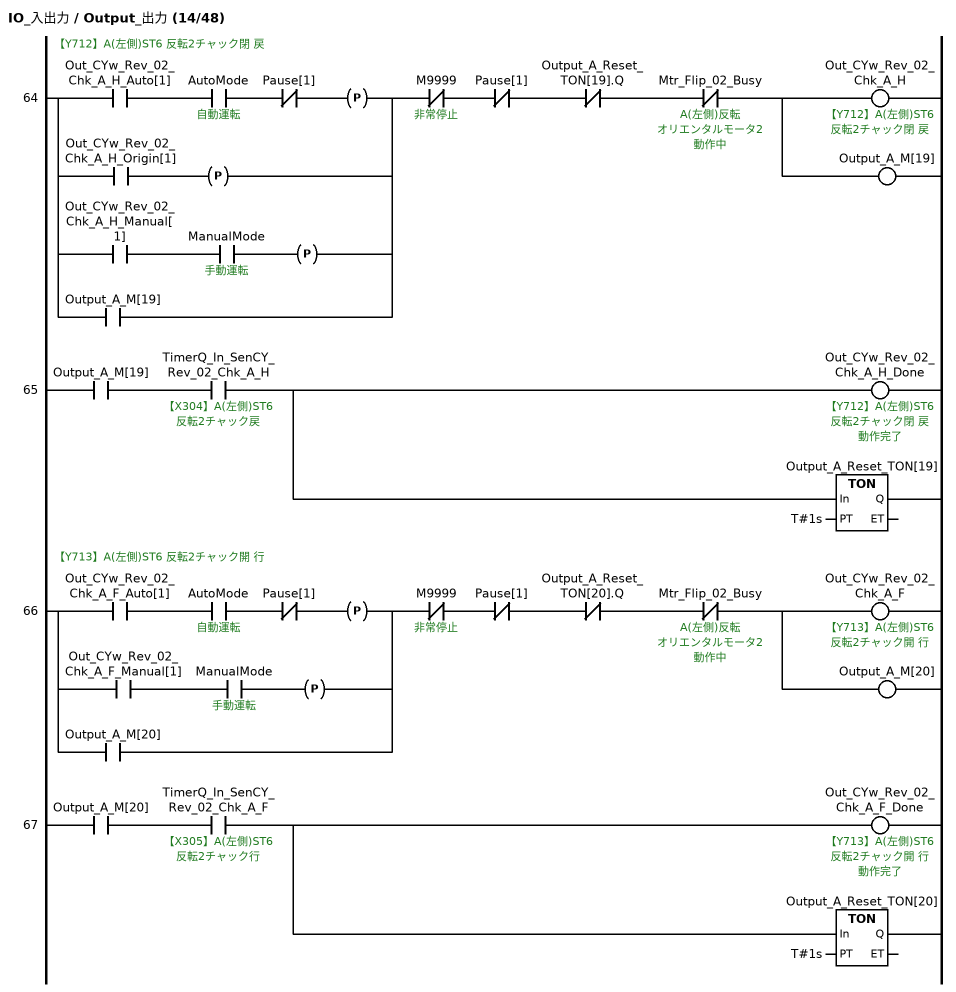
(* Rung 64: 【Y712】A(左側)ST6 反転2チャック閉 戻 *)
_e83(CLK := Out_CYw_Rev_02_Chk_A_H_Auto[1] AND AutoMode AND NOT Pause[1]);
_e84(CLK := Out_CYw_Rev_02_Chk_A_H_Origin[1]);
_e85(CLK := Out_CYw_Rev_02_Chk_A_H_Manual[1] AND ManualMode);
_p86 := (_e83.Q OR _e84.Q OR _e85.Q OR Output_A_M[19]) AND NOT M9999 AND NOT Pause[1] AND NOT Output_A_Reset_TON[19].Q AND NOT Mtr_Flip_02_Busy;
Out_CYw_Rev_02_Chk_A_H := _p86;
Output_A_M[19] := _p86;
(* Rung 65 *)
_p87 := Output_A_M[19] AND TimerQ_In_SenCY_Rev_02_Chk_A_H;
Out_CYw_Rev_02_Chk_A_H_Done := _p87;
Output_A_Reset_TON[19](In := _p87, PT := T#1s);
(* Rung 66: 【Y713】A(左側)ST6 反転2チャック開 行 *)
_e88(CLK := Out_CYw_Rev_02_Chk_A_F_Auto[1] AND AutoMode AND NOT Pause[1]);
_e89(CLK := Out_CYw_Rev_02_Chk_A_F_Manual[1] AND ManualMode);
_p90 := (_e88.Q OR _e89.Q OR Output_A_M[20]) AND NOT M9999 AND NOT Pause[1] AND NOT Output_A_Reset_TON[20].Q AND NOT Mtr_Flip_02_Busy;
Out_CYw_Rev_02_Chk_A_F := _p90;
Output_A_M[20] := _p90;
(* Rung 67 *)
_p91 := Output_A_M[20] AND TimerQ_In_SenCY_Rev_02_Chk_A_F;
Out_CYw_Rev_02_Chk_A_F_Done := _p91;
Output_A_Reset_TON[20](In := _p91, PT := T#1s);

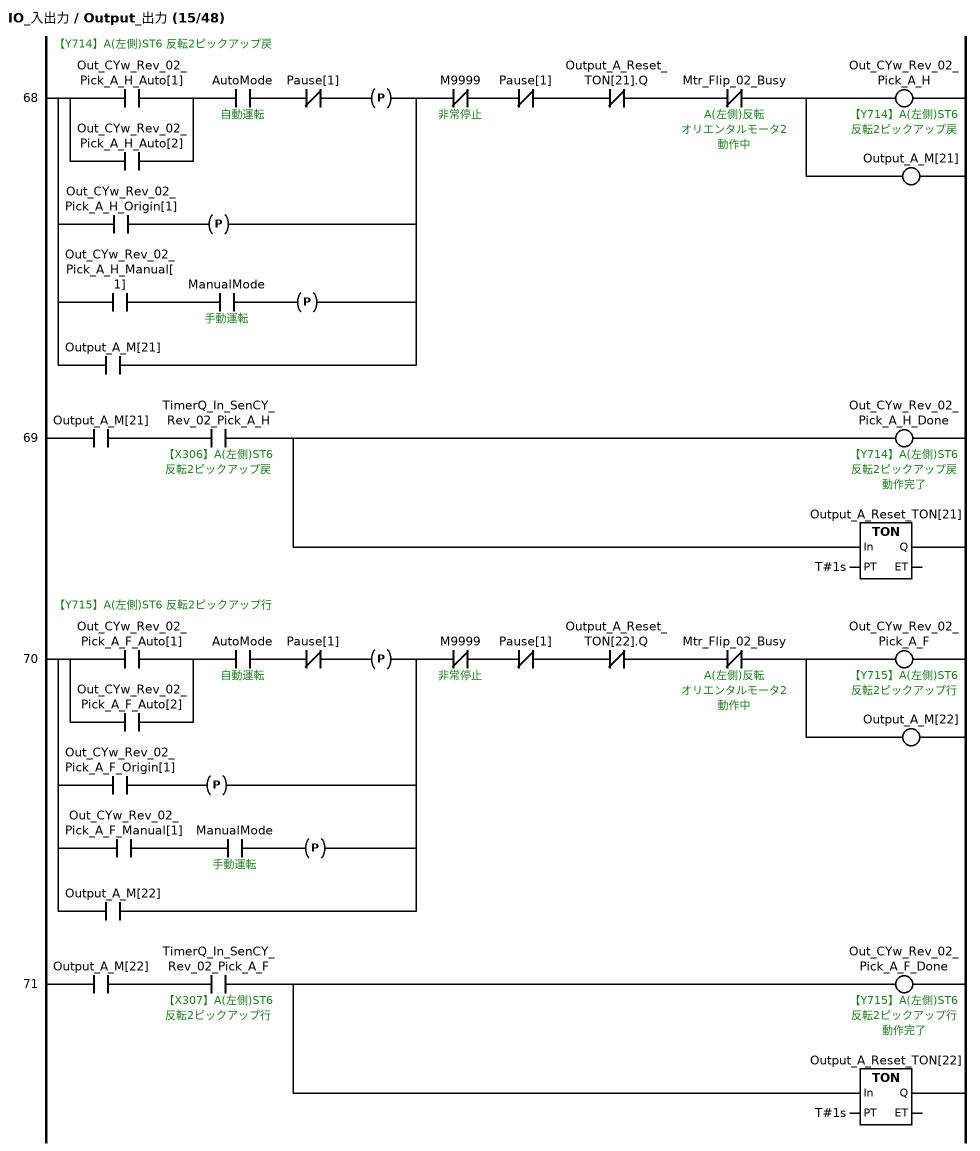
(* Rung 68: 【Y714】A(左側)ST6 反転2ピックアップ戻 *)
_e92(CLK := (Out_CYw_Rev_02_Pick_A_H_Auto[1] OR Out_CYw_Rev_02_Pick_A_H_Auto[2]) AND AutoMode AND NOT Pause[1]);
_e93(CLK := Out_CYw_Rev_02_Pick_A_H_Origin[1]);
_e94(CLK := Out_CYw_Rev_02_Pick_A_H_Manual[1] AND ManualMode);
_p95 := (_e92.Q OR _e93.Q OR _e94.Q OR Output_A_M[21]) AND NOT M9999 AND NOT Pause[1] AND NOT Output_A_Reset_TON[21].Q AND NOT Mtr_Flip_02_Busy;
Out_CYw_Rev_02_Pick_A_H := _p95;
Output_A_M[21] := _p95;
(* Rung 69 *)
_p96 := Output_A_M[21] AND TimerQ_In_SenCY_Rev_02_Pick_A_H;
Out_CYw_Rev_02_Pick_A_H_Done := _p96;
Output_A_Reset_TON[21](In := _p96, PT := T#1s);
(* Rung 70: 【Y715】A(左側)ST6 反転2ピックアップ行 *)
_e97(CLK := (Out_CYw_Rev_02_Pick_A_F_Auto[1] OR Out_CYw_Rev_02_Pick_A_F_Auto[2]) AND AutoMode AND NOT Pause[1]);
_e98(CLK := Out_CYw_Rev_02_Pick_A_F_Origin[1]);
_e99(CLK := Out_CYw_Rev_02_Pick_A_F_Manual[1] AND ManualMode);
_p100 := (_e97.Q OR _e98.Q OR _e99.Q OR Output_A_M[22]) AND NOT M9999 AND NOT Pause[1] AND NOT Output_A_Reset_TON[22].Q AND NOT Mtr_Flip_02_Busy;
Out_CYw_Rev_02_Pick_A_F := _p100;
Output_A_M[22] := _p100;
(* Rung 71 *)
_p101 := Output_A_M[22] AND TimerQ_In_SenCY_Rev_02_Pick_A_F;
Out_CYw_Rev_02_Pick_A_F_Done := _p101;
Output_A_Reset_TON[22](In := _p101, PT := T#1s);

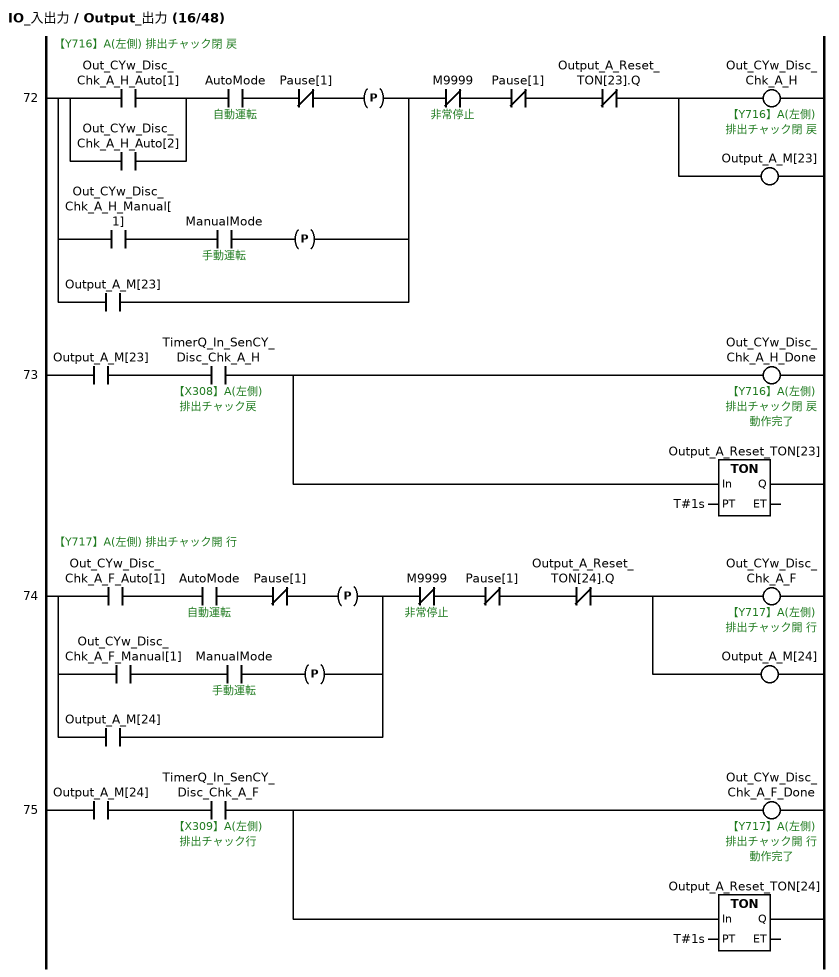
(* Rung 72: 【Y716】A(左側) 排出チャック閉 戻 *)
_e102(CLK := (Out_CYw_Disc_Chk_A_H_Auto[1] OR Out_CYw_Disc_Chk_A_H_Auto[2]) AND AutoMode AND NOT Pause[1]);
_e103(CLK := Out_CYw_Disc_Chk_A_H_Manual[1] AND ManualMode);
_p104 := (_e102.Q OR _e103.Q OR Output_A_M[23]) AND NOT M9999 AND NOT Pause[1] AND NOT Output_A_Reset_TON[23].Q;
Out_CYw_Disc_Chk_A_H := _p104;
Output_A_M[23] := _p104;
(* Rung 73 *)
Out_CYw_Disc_Chk_A_H_Done := Output_A_M[23] AND TimerQ_In_SenCY_Disc_Chk_A_H;
Output_A_Reset_TON[23](In := Output_A_M[23] AND TimerQ_In_SenCY_Disc_Chk_A_H, PT := T#1s);
(* Rung 74: 【Y717】A(左側) 排出チャック開 行 *)
_e105(CLK := Out_CYw_Disc_Chk_A_F_Auto[1] AND AutoMode AND NOT Pause[1]);
_e106(CLK := Out_CYw_Disc_Chk_A_F_Manual[1] AND ManualMode);
_p107 := (_e105.Q OR _e106.Q OR Output_A_M[24]) AND NOT M9999 AND NOT Pause[1] AND NOT Output_A_Reset_TON[24].Q;
Out_CYw_Disc_Chk_A_F := _p107;
Output_A_M[24] := _p107;
(* Rung 75 *)
Out_CYw_Disc_Chk_A_F_Done := Output_A_M[24] AND TimerQ_In_SenCY_Disc_Chk_A_F;
Output_A_Reset_TON[24](In := Output_A_M[24] AND TimerQ_In_SenCY_Disc_Chk_A_F, PT := T#1s);

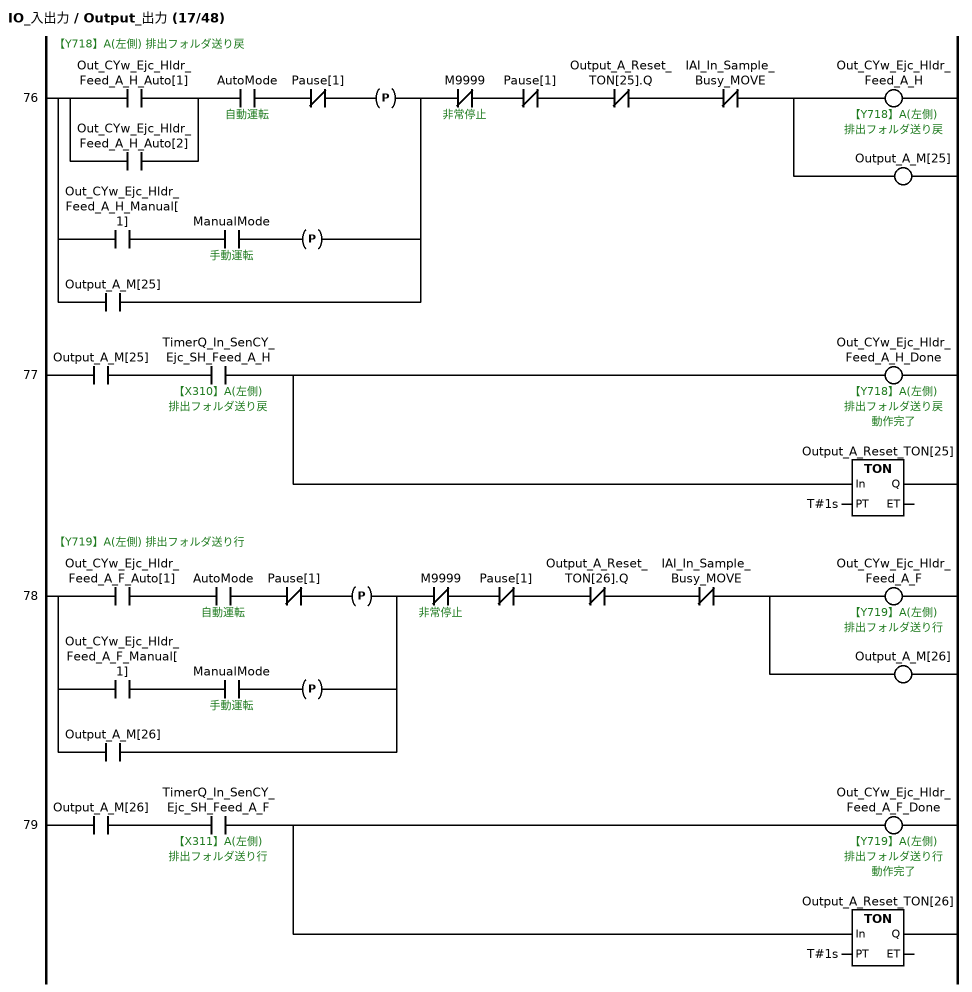
(* Rung 76: 【Y718】A(左側) 排出フォルダ送り戻 *)
_e108(CLK := (Out_CYw_Ejc_Hldr_Feed_A_H_Auto[1] OR Out_CYw_Ejc_Hldr_Feed_A_H_Auto[2]) AND AutoMode AND NOT Pause[1]);
_e109(CLK := Out_CYw_Ejc_Hldr_Feed_A_H_Manual[1] AND ManualMode);
_p110 := (_e108.Q OR _e109.Q OR Output_A_M[25]) AND NOT M9999 AND NOT Pause[1] AND NOT Output_A_Reset_TON[25].Q AND NOT IAI_In_Sample_Busy_MOVE;
Out_CYw_Ejc_Hldr_Feed_A_H := _p110;
Output_A_M[25] := _p110;
(* Rung 77 *)
_p111 := Output_A_M[25] AND TimerQ_In_SenCY_Ejc_SH_Feed_A_H;
Out_CYw_Ejc_Hldr_Feed_A_H_Done := _p111;
Output_A_Reset_TON[25](In := _p111, PT := T#1s);
(* Rung 78: 【Y719】A(左側) 排出フォルダ送り行 *)
_e112(CLK := Out_CYw_Ejc_Hldr_Feed_A_F_Auto[1] AND AutoMode AND NOT Pause[1]);
_e113(CLK := Out_CYw_Ejc_Hldr_Feed_A_F_Manual[1] AND ManualMode);
_p114 := (_e112.Q OR _e113.Q OR Output_A_M[26]) AND NOT M9999 AND NOT Pause[1] AND NOT Output_A_Reset_TON[26].Q AND NOT IAI_In_Sample_Busy_MOVE;
Out_CYw_Ejc_Hldr_Feed_A_F := _p114;
Output_A_M[26] := _p114;
(* Rung 79 *)
_p115 := Output_A_M[26] AND TimerQ_In_SenCY_Ejc_SH_Feed_A_F;
Out_CYw_Ejc_Hldr_Feed_A_F_Done := _p115;
Output_A_Reset_TON[26](In := _p115, PT := T#1s);

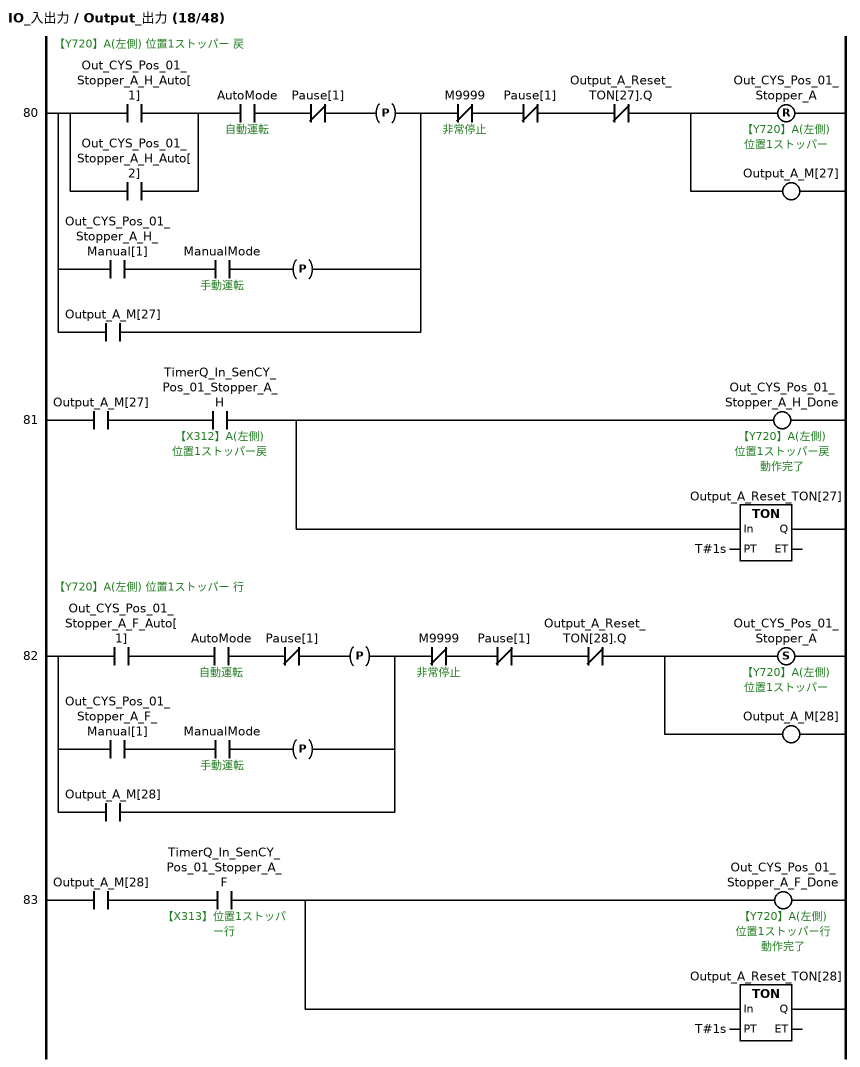
(* Rung 80: 【Y720】A(左側) 位置1ストッパー 戻 *)
_e116(CLK := (Out_CYS_Pos_01_Stopper_A_H_Auto[1] OR Out_CYS_Pos_01_Stopper_A_H_Auto[2]) AND AutoMode AND NOT Pause[1]);
_e117(CLK := Out_CYS_Pos_01_Stopper_A_H_Manual[1] AND ManualMode);
_p118 := (_e116.Q OR _e117.Q OR Output_A_M[27]) AND NOT M9999 AND NOT Pause[1] AND NOT Output_A_Reset_TON[27].Q;
IF _p118 THEN Out_CYS_Pos_01_Stopper_A := FALSE; END_IF;
Output_A_M[27] := _p118;
(* Rung 81 *)
_p119 := Output_A_M[27] AND TimerQ_In_SenCY_Pos_01_Stopper_A_H;
Out_CYS_Pos_01_Stopper_A_H_Done := _p119;
Output_A_Reset_TON[27](In := _p119, PT := T#1s);
(* Rung 82: 【Y720】A(左側) 位置1ストッパー 行 *)
_e120(CLK := Out_CYS_Pos_01_Stopper_A_F_Auto[1] AND AutoMode AND NOT Pause[1]);
_e121(CLK := Out_CYS_Pos_01_Stopper_A_F_Manual[1] AND ManualMode);
_p122 := (_e120.Q OR _e121.Q OR Output_A_M[28]) AND NOT M9999 AND NOT Pause[1] AND NOT Output_A_Reset_TON[28].Q;
IF _p122 THEN Out_CYS_Pos_01_Stopper_A := TRUE; END_IF;
Output_A_M[28] := _p122;
(* Rung 83 *)
_p123 := Output_A_M[28] AND TimerQ_In_SenCY_Pos_01_Stopper_A_F;
Out_CYS_Pos_01_Stopper_A_F_Done := _p123;
Output_A_Reset_TON[28](In := _p123, PT := T#1s);

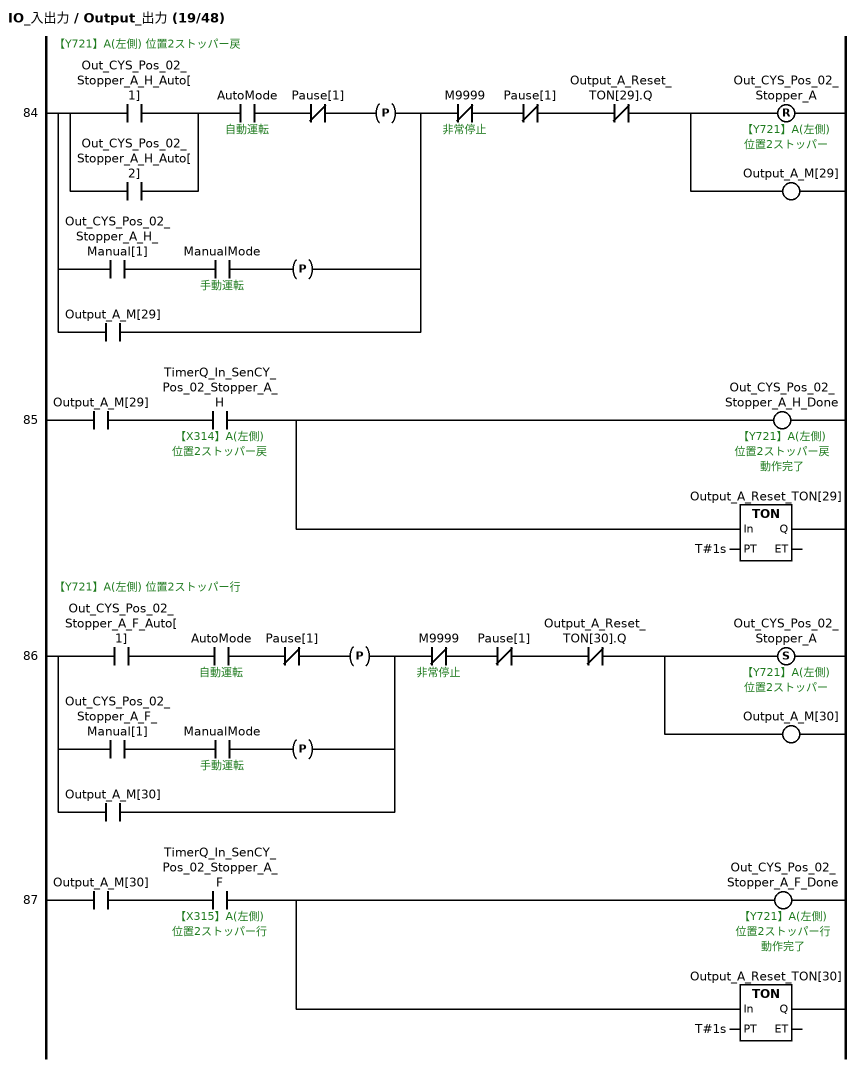
(* Rung 84: 【Y721】A(左側) 位置2ストッパー戻 *)
_e124(CLK := (Out_CYS_Pos_02_Stopper_A_H_Auto[1] OR Out_CYS_Pos_02_Stopper_A_H_Auto[2]) AND AutoMode AND NOT Pause[1]);
_e125(CLK := Out_CYS_Pos_02_Stopper_A_H_Manual[1] AND ManualMode);
_p126 := (_e124.Q OR _e125.Q OR Output_A_M[29]) AND NOT M9999 AND NOT Pause[1] AND NOT Output_A_Reset_TON[29].Q;
IF _p126 THEN Out_CYS_Pos_02_Stopper_A := FALSE; END_IF;
Output_A_M[29] := _p126;
(* Rung 85 *)
_p127 := Output_A_M[29] AND TimerQ_In_SenCY_Pos_02_Stopper_A_H;
Out_CYS_Pos_02_Stopper_A_H_Done := _p127;
Output_A_Reset_TON[29](In := _p127, PT := T#1s);
(* Rung 86: 【Y721】A(左側) 位置2ストッパー行 *)
_e128(CLK := Out_CYS_Pos_02_Stopper_A_F_Auto[1] AND AutoMode AND NOT Pause[1]);
_e129(CLK := Out_CYS_Pos_02_Stopper_A_F_Manual[1] AND ManualMode);
_p130 := (_e128.Q OR _e129.Q OR Output_A_M[30]) AND NOT M9999 AND NOT Pause[1] AND NOT Output_A_Reset_TON[30].Q;
IF _p130 THEN Out_CYS_Pos_02_Stopper_A := TRUE; END_IF;
Output_A_M[30] := _p130;
(* Rung 87 *)
_p131 := Output_A_M[30] AND TimerQ_In_SenCY_Pos_02_Stopper_A_F;
Out_CYS_Pos_02_Stopper_A_F_Done := _p131;
Output_A_Reset_TON[30](In := _p131, PT := T#1s);

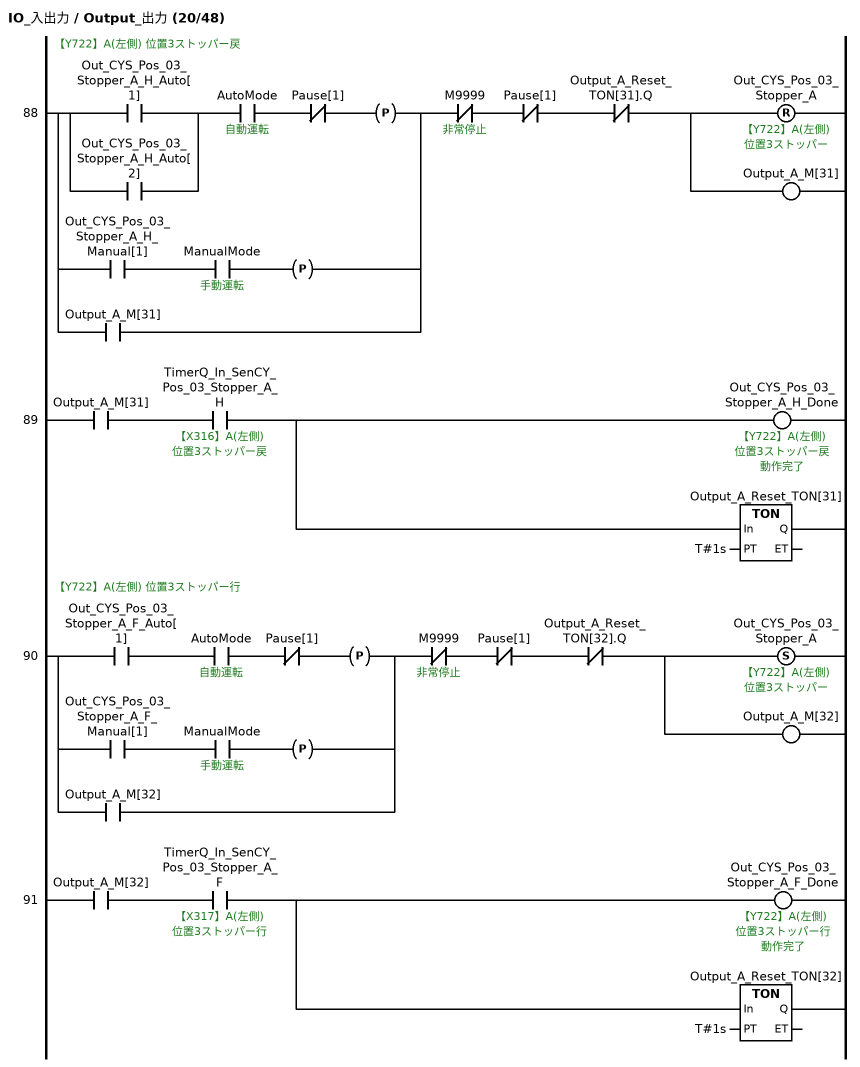
(* Rung 88: 【Y722】A(左側) 位置3ストッパー戻 *)
_e132(CLK := (Out_CYS_Pos_03_Stopper_A_H_Auto[1] OR Out_CYS_Pos_03_Stopper_A_H_Auto[2]) AND AutoMode AND NOT Pause[1]);
_e133(CLK := Out_CYS_Pos_03_Stopper_A_H_Manual[1] AND ManualMode);
_p134 := (_e132.Q OR _e133.Q OR Output_A_M[31]) AND NOT M9999 AND NOT Pause[1] AND NOT Output_A_Reset_TON[31].Q;
IF _p134 THEN Out_CYS_Pos_03_Stopper_A := FALSE; END_IF;
Output_A_M[31] := _p134;
(* Rung 89 *)
_p135 := Output_A_M[31] AND TimerQ_In_SenCY_Pos_03_Stopper_A_H;
Out_CYS_Pos_03_Stopper_A_H_Done := _p135;
Output_A_Reset_TON[31](In := _p135, PT := T#1s);
(* Rung 90: 【Y722】A(左側) 位置3ストッパー行 *)
_e136(CLK := Out_CYS_Pos_03_Stopper_A_F_Auto[1] AND AutoMode AND NOT Pause[1]);
_e137(CLK := Out_CYS_Pos_03_Stopper_A_F_Manual[1] AND ManualMode);
_p138 := (_e136.Q OR _e137.Q OR Output_A_M[32]) AND NOT M9999 AND NOT Pause[1] AND NOT Output_A_Reset_TON[32].Q;
IF _p138 THEN Out_CYS_Pos_03_Stopper_A := TRUE; END_IF;
Output_A_M[32] := _p138;
(* Rung 91 *)
_p139 := Output_A_M[32] AND TimerQ_In_SenCY_Pos_03_Stopper_A_F;
Out_CYS_Pos_03_Stopper_A_F_Done := _p139;
Output_A_Reset_TON[32](In := _p139, PT := T#1s);

